FUNCTION_BLOCK "Conveyor_HMI_FB_1"   // FB 13, author

VAR_INPUT
   HMI_No : UInt;
   Sys_No : UInt;
   Zone : UInt;
END_VAR

VAR_IN_OUT
   Enable : Bool;
   Mode_Change : UInt;
   Transfer_To_ID : DInt;
   Transfer_From_ID : DInt;
   Pallet_Allignment : Bool;
   Enable(1) : Bool;
   Mode_Change(1) : UInt;
   Transfer_To_ID(1) : DInt;
   Transfer_From_ID(1) : DInt;
   Pallet_Allignment(1) : Bool;
END_VAR

VAR
   R_Charge_Cnv_Commands : R_TRIG;
   T_Reset_Charge : TON_TIME;
   ID : DInt;
   ID(1) : DInt;
   ID_Old : DInt;
   ID_Old(1) : DInt;
END_VAR

VAR_TEMP
   i : UInt;
   J : UInt;
   No_Light_Guard : Bool;
END_VAR

BEGIN
CNV_Selector_1(Sys_No := #Sys_No,
                 Zone:= #Zone,
                 CNV1_2_Selected := "CNV_HMI".CNV2_Selected[#HMI_No],
                 ID => #ID,
                 ID(1) => #"ID(1)");


REGION SEND/RECEIVE BUTTON
    IF NOT "Control_DB".VTD_Sys[#Sys_No].Running AND "Control_DB".VTD_Sys[#Sys_No].Current_Level <> 0 THEN
        IF "CNV_HMI".CNV2_Selected[#HMI_No] = 1 AND "HMI_DB".ScreenNo[#HMI_No] = 2 THEN
            //CNV 1
            IF "Control_DB".ECnv_Sys[#Sys_No].Cnv_Occupied AND NOT "Control_DB".LCnv_Sys[#Sys_No].Cnv_Level["Control_DB".VTD_Sys[#Sys_No].Current_Level].Cnv1.Cnv_Occupied AND
                NOT "Control_DB".ECnv_Sys[#Sys_No].Running AND NOT "Control_DB".LCnv_Sys[#Sys_No].Cnv_Level["Control_DB".VTD_Sys[#Sys_No].Current_Level].Cnv1.Running THEN
                "CNV_HMI".In_Out[#HMI_No] := TRUE;
            ELSIF NOT "Control_DB".ECnv_Sys[#Sys_No].Cnv_Occupied AND "Control_DB".LCnv_Sys[#Sys_No].Cnv_Level["Control_DB".VTD_Sys[#Sys_No].Current_Level].Cnv1.Cnv_Occupied AND
                NOT "Control_DB".ECnv_Sys[#Sys_No].Running AND NOT "Control_DB".LCnv_Sys[#Sys_No].Cnv_Level["Control_DB".VTD_Sys[#Sys_No].Current_Level].Cnv1.Running THEN
                "CNV_HMI".In_Out[#HMI_No] := FALSE;
            ELSE
                ;
            END_IF;
            //CNV 2
        ELSIF "CNV_HMI".CNV2_Selected[#HMI_No] = 2 AND "HMI_DB".ScreenNo[#HMI_No] = 2 THEN   //CNV 2
            IF "Control_DB".ECnv_Sys[#Sys_No].Cnv_Occupied AND NOT "Control_DB".LCnv_Sys[#Sys_No].Cnv_Level["Control_DB".VTD_Sys[#Sys_No].Current_Level].Cnv2.Cnv_Occupied AND
                NOT "Control_DB".ECnv_Sys[#Sys_No].Running AND NOT "Control_DB".LCnv_Sys[#Sys_No].Cnv_Level["Control_DB".VTD_Sys[#Sys_No].Current_Level].Cnv2.Running THEN
                "CNV_HMI".In_Out[#HMI_No] := TRUE;
            ELSIF NOT "Control_DB".ECnv_Sys[#Sys_No].Cnv_Occupied AND "Control_DB".LCnv_Sys[#Sys_No].Cnv_Level["Control_DB".VTD_Sys[#Sys_No].Current_Level].Cnv2.Cnv_Occupied AND
                NOT "Control_DB".ECnv_Sys[#Sys_No].Running AND NOT "Control_DB".LCnv_Sys[#Sys_No].Cnv_Level["Control_DB".VTD_Sys[#Sys_No].Current_Level].Cnv2.Running THEN
                "CNV_HMI".In_Out[#HMI_No] := FALSE;
            ELSE
                ;
            END_IF;
        END_IF;
    END_IF;
END_REGION ;

REGION Assign Conveyor 1
    REGION CHARGE DATA FROM THE CORRECT CONVEYOR
        //CHARGE DATA CHANGING CONVEYORS ID
        IF #ID <> #ID_Old THEN
            "CNV_HMI".Charge_Commands[#HMI_No] := TRUE;
            #ID_Old := #ID;
        END_IF;
        #R_Charge_Cnv_Commands();

        #R_Charge_Cnv_Commands(CLK := "CNV_HMI".Charge_Commands[#HMI_No]);

        //CHARGE ONCE THE COMMANDS
        IF "CNV_HMI".Charge_Commands[#Sys_No] THEN
            #Enable := "Control_DB".ECnv_Sys[#Sys_No].Instruction.Enable;
            #Mode_Change := "Control_DB".ECnv_Sys[#Sys_No].Instruction.Mode_Change;
            #Transfer_To_ID := "Control_DB".ECnv_Sys[#Sys_No].Instruction.Transfer_To_ID;
            #Transfer_From_ID := "Control_DB".ECnv_Sys[#Sys_No].Instruction.Transfer_From_ID;
            #Pallet_Allignment := "Control_DB".ECnv_Sys[#Sys_No].Instruction.Pallet_Allignment;
        END_IF;
    END_REGION

    REGION CHARGE DATA FROM HMI (AFTER CHARGE DATA)
        IF NOT "CNV_HMI".Charge_Commands[#HMI_No] AND NOT #R_Charge_Cnv_Commands.Q THEN
            CASE #ID OF
                    //SYSTEM 1
                120101:
                    Feed_ECNV_1(HMI_No := #HMI_No,
                                  HMI_Box:= #Zone,
                                  Overhang_Left:="CVTD1 OVERHANG LEFT",
                                  Overhang_Right:="CVTD1 OVERHANG RIGHT",
                                  Sys_No := #Sys_No,
                                  Safety_OK := "Remote_Panel_DB_1".Safety_OK);
                120201:
                    Feed_ECNV_1(HMI_No := #HMI_No,
                                  HMI_Box:= #Zone,
                                  Overhang_Left:="CVTD1 OVERHANG LEFT",
                                  Overhang_Right:="CVTD1 OVERHANG RIGHT",
                                  Sys_No := #Sys_No,
                                  Safety_OK := "Remote_Panel_DB_1".Safety_OK);
                120301:
                    Feed_ECNV_1(HMI_No := #HMI_No,
                                  HMI_Box:= #Zone,
                                  Overhang_Left:="CVTD1 OVERHANG LEFT",
                                  Overhang_Right:="CVTD1 OVERHANG RIGHT",
                                  Sys_No := #Sys_No,
                                  Safety_OK := "Remote_Panel_DB_1".Safety_OK);
                120401:
                    Feed_ECNV_1(HMI_No := #HMI_No,
                                  HMI_Box:= #Zone,
                                  Overhang_Left:="CVTD1 OVERHANG LEFT",
                                  Overhang_Right:="CVTD1 OVERHANG RIGHT",
                                  Sys_No := #Sys_No,
                                  Safety_OK := "Remote_Panel_DB_1".Safety_OK);
                120501:
                    Feed_ECNV_1(HMI_No := #HMI_No,
                                  HMI_Box:= #Zone,
                                  Overhang_Left:="CVTD1 OVERHANG LEFT",
                                  Overhang_Right:="CVTD1 OVERHANG RIGHT",
                                  Sys_No := #Sys_No,
                                  Safety_OK := "Remote_Panel_DB_1".Safety_OK);
                120601:
                    Feed_ECNV_1(HMI_No := #HMI_No,
                                  HMI_Box:= #Zone,
                                  Overhang_Left:="CVTD1 OVERHANG LEFT",
                                  Overhang_Right:="CVTD1 OVERHANG RIGHT",
                                  Sys_No := #Sys_No,
                                  Safety_OK := "Remote_Panel_DB_1".Safety_OK);
                120701:
                    Feed_ECNV_1(HMI_No := #HMI_No,
                                  HMI_Box:= #Zone,
                                  Overhang_Left:="CVTD1 OVERHANG LEFT",
                                  Overhang_Right:="CVTD1 OVERHANG RIGHT",
                                  Sys_No := #Sys_No,
                                  Safety_OK := "Remote_Panel_DB_1".Safety_OK);
                120801:
                    Feed_ECNV_1(HMI_No := #HMI_No,
                                  HMI_Box:= #Zone,
                                  Overhang_Left:="CVTD1 OVERHANG LEFT",
                                  Overhang_Right:="CVTD1 OVERHANG RIGHT",
                                  Sys_No := #Sys_No,
                                  Safety_OK := "Remote_Panel_DB_1".Safety_OK);

                    //SYSTEM 2
                120102:
                    Feed_ECNV_1(HMI_No := #HMI_No,
                                  HMI_Box:= #Zone,
                                  Overhang_Left:="CVTD2 OVERHANG LEFT",
                                  Overhang_Right:="CVTD2 OVERHANG RIGHT",
                                  Sys_No := 2,
                                  Safety_OK := "Remote_Panel_DB_2".Safety_OK);
                120202:
                    Feed_ECNV_1(HMI_No := #HMI_No,
                                  HMI_Box:= #Zone,
                                  Overhang_Left:="CVTD2 OVERHANG LEFT",
                                  Overhang_Right:="CVTD2 OVERHANG RIGHT",
                                  Sys_No := 2,
                                  Safety_OK := "Remote_Panel_DB_2".Safety_OK);
                120302:
                    Feed_ECNV_1(HMI_No := #HMI_No,
                                  HMI_Box:= #Zone,
                                  Overhang_Left:="CVTD2 OVERHANG LEFT",
                                  Overhang_Right:="CVTD2 OVERHANG RIGHT",
                                  Sys_No := 2,
                                  Safety_OK := "Remote_Panel_DB_2".Safety_OK);
                120402:
                    Feed_ECNV_1(HMI_No := #HMI_No,
                                  HMI_Box:= #Zone,
                                  Overhang_Left:="CVTD2 OVERHANG LEFT",
                                  Overhang_Right:="CVTD2 OVERHANG RIGHT",
                                  Sys_No := 2,
                                  Safety_OK := "Remote_Panel_DB_2".Safety_OK);
                120502:
                    Feed_ECNV_1(HMI_No := #HMI_No,
                                  HMI_Box:= #Zone,
                                  Overhang_Left:="CVTD2 OVERHANG LEFT",
                                  Overhang_Right:="CVTD2 OVERHANG RIGHT",
                                  Sys_No := 2,
                                  Safety_OK := "Remote_Panel_DB_2".Safety_OK);
                120602:
                    Feed_ECNV_1(HMI_No := #HMI_No,
                                  HMI_Box:= #Zone,
                                  Overhang_Left:="CVTD2 OVERHANG LEFT",
                                  Overhang_Right:="CVTD2 OVERHANG RIGHT",
                                  Sys_No := 2,
                                  Safety_OK := "Remote_Panel_DB_2".Safety_OK);
                120702:
                    Feed_ECNV_1(HMI_No := #HMI_No,
                                  HMI_Box:= #Zone,
                                  Overhang_Left:="CVTD2 OVERHANG LEFT",
                                  Overhang_Right:="CVTD2 OVERHANG RIGHT",
                                  Sys_No := 2,
                                  Safety_OK := "Remote_Panel_DB_2".Safety_OK);
                120802:
                    Feed_ECNV_1(HMI_No := #HMI_No,
                                  HMI_Box:= #Zone,
                                  Overhang_Left:="CVTD2 OVERHANG LEFT",
                                  Overhang_Right:="CVTD2 OVERHANG RIGHT",
                                  Sys_No := 2,
                                  Safety_OK := "Remote_Panel_DB_2".Safety_OK);

                    //SYSTEM 3
                120103:
                    Feed_ECNV_1(HMI_No := #HMI_No,
                                  HMI_Box:= #Zone,
                                  Overhang_Left:="CVTD3 OVERHANG LEFT",
                                  Overhang_Right:="CVTD3 OVERHANG RIGHT",
                                  Sys_No := 3,
                                  Safety_OK := "Remote_Panel_DB_3".Safety_OK);
                120203:
                    Feed_ECNV_1(HMI_No := #HMI_No,
                                  HMI_Box:= #Zone,
                                  Overhang_Left:="CVTD3 OVERHANG LEFT",
                                  Overhang_Right:="CVTD3 OVERHANG RIGHT",
                                  Sys_No := 3,
                                  Safety_OK := "Remote_Panel_DB_3".Safety_OK);
                120303:
                    Feed_ECNV_1(HMI_No := #HMI_No,
                                  HMI_Box:= #Zone,
                                  Overhang_Left:="CVTD3 OVERHANG LEFT",
                                  Overhang_Right:="CVTD3 OVERHANG RIGHT",
                                  Sys_No := 3,
                                  Safety_OK := "Remote_Panel_DB_3".Safety_OK);
                120403:
                    Feed_ECNV_1(HMI_No := #HMI_No,
                                  HMI_Box:= #Zone,
                                  Overhang_Left:="CVTD3 OVERHANG LEFT",
                                  Overhang_Right:="CVTD3 OVERHANG RIGHT",
                                  Sys_No := 3,
                                  Safety_OK := "Remote_Panel_DB_3".Safety_OK);
                120503:
                    Feed_ECNV_1(HMI_No := #HMI_No,
                                  HMI_Box:= #Zone,
                                  Overhang_Left:="CVTD3 OVERHANG LEFT",
                                  Overhang_Right:="CVTD3 OVERHANG RIGHT",
                                  Sys_No := 3,
                                  Safety_OK := "Remote_Panel_DB_3".Safety_OK);
                120603:
                    Feed_ECNV_1(HMI_No := #HMI_No,
                                  HMI_Box:= #Zone,
                                  Overhang_Left:="CVTD3 OVERHANG LEFT",
                                  Overhang_Right:="CVTD3 OVERHANG RIGHT",
                                  Sys_No := 3,
                                  Safety_OK := "Remote_Panel_DB_3".Safety_OK);
                120703:
                    Feed_ECNV_1(HMI_No := #HMI_No,
                                  HMI_Box:= #Zone,
                                  Overhang_Left:="CVTD3 OVERHANG LEFT",
                                  Overhang_Right:="CVTD3 OVERHANG RIGHT",
                                  Sys_No := 3,
                                  Safety_OK := "Remote_Panel_DB_3".Safety_OK);
                120803:
                    Feed_ECNV_1(HMI_No := #HMI_No,
                                  HMI_Box:= #Zone,
                                  Overhang_Left:="CVTD3 OVERHANG LEFT",
                                  Overhang_Right:="CVTD3 OVERHANG RIGHT",
                                  Sys_No := 3,
                                  Safety_OK := "Remote_Panel_DB_3".Safety_OK);

                    //SYSTEM 4
                120104:
                    Feed_ECNV_1(HMI_No := #HMI_No,
                                  HMI_Box:= #Zone,
                                  Overhang_Left:="CVTD4 OVERHANG LEFT",
                                  Overhang_Right:="CVTD4 OVERHANG RIGHT",
                                  Sys_No := 4,
                                  Safety_OK := "Remote_Panel_DB_4".Safety_OK);
                120204:
                    Feed_ECNV_1(HMI_No := #HMI_No,
                                  HMI_Box:= #Zone,
                                  Overhang_Left:="CVTD4 OVERHANG LEFT",
                                  Overhang_Right:="CVTD4 OVERHANG RIGHT",
                                  Sys_No := 4,
                                  Safety_OK := "Remote_Panel_DB_4".Safety_OK);
                120304:
                    Feed_ECNV_1(HMI_No := #HMI_No,
                                  HMI_Box:= #Zone,
                                  Overhang_Left:="CVTD4 OVERHANG LEFT",
                                  Overhang_Right:="CVTD4 OVERHANG RIGHT",
                                  Sys_No := 4,
                                  Safety_OK := "Remote_Panel_DB_4".Safety_OK);
                120404:
                    Feed_ECNV_1(HMI_No := #HMI_No,
                                  HMI_Box:= #Zone,
                                  Overhang_Left:="CVTD4 OVERHANG LEFT",
                                  Overhang_Right:="CVTD4 OVERHANG RIGHT",
                                  Sys_No := 4,
                                  Safety_OK := "Remote_Panel_DB_4".Safety_OK);
                120504:
                    Feed_ECNV_1(HMI_No := #HMI_No,
                                  HMI_Box:= #Zone,
                                  Overhang_Left:="CVTD4 OVERHANG LEFT",
                                  Overhang_Right:="CVTD4 OVERHANG RIGHT",
                                  Sys_No := 4,
                                  Safety_OK := "Remote_Panel_DB_4".Safety_OK);
                120604:
                    Feed_ECNV_1(HMI_No := #HMI_No,
                                  HMI_Box:= #Zone,
                                  Overhang_Left:="CVTD4 OVERHANG LEFT",
                                  Overhang_Right:="CVTD4 OVERHANG RIGHT",
                                  Sys_No := 4,
                                  Safety_OK := "Remote_Panel_DB_4".Safety_OK);
                120704:
                    Feed_ECNV_1(HMI_No := #HMI_No,
                                  HMI_Box:= #Zone,
                                  Overhang_Left:="CVTD4 OVERHANG LEFT",
                                  Overhang_Right:="CVTD4 OVERHANG RIGHT",
                                  Sys_No := 4,
                                  Safety_OK := "Remote_Panel_DB_4".Safety_OK);
                120804:
                    Feed_ECNV_1(HMI_No := #HMI_No,
                                  HMI_Box:= #Zone,
                                  Overhang_Left:="CVTD4 OVERHANG LEFT",
                                  Overhang_Right:="CVTD4 OVERHANG RIGHT",
                                  Sys_No := 4,
                                  Safety_OK := "Remote_Panel_DB_4".Safety_OK);

                    //SYSTEM 5
                120105:
                    Feed_ECNV_1(HMI_No := #HMI_No,
                                  HMI_Box:= #Zone,
                                  Overhang_Left:="CVTD5 OVERHANG LEFT",
                                  Overhang_Right:="CVTD5 OVERHANG RIGHT",
                                  Sys_No := 5,
                                  Safety_OK := "Remote_Panel_DB_5".Safety_OK);
                120205:
                    Feed_ECNV_1(HMI_No := #HMI_No,
                                  HMI_Box:= #Zone,
                                  Overhang_Left:="CVTD5 OVERHANG LEFT",
                                  Overhang_Right:="CVTD5 OVERHANG RIGHT",
                                  Sys_No := 5,
                                  Safety_OK := "Remote_Panel_DB_5".Safety_OK);
                120305:
                    Feed_ECNV_1(HMI_No := #HMI_No,
                                  HMI_Box:= #Zone,
                                  Overhang_Left:="CVTD5 OVERHANG LEFT",
                                  Overhang_Right:="CVTD5 OVERHANG RIGHT",
                                  Sys_No := 5,
                                  Safety_OK := "Remote_Panel_DB_5".Safety_OK);
                120405:
                    Feed_ECNV_1(HMI_No := #HMI_No,
                                  HMI_Box:= #Zone,
                                  Overhang_Left:="CVTD5 OVERHANG LEFT",
                                  Overhang_Right:="CVTD5 OVERHANG RIGHT",
                                  Sys_No := 5,
                                  Safety_OK := "Remote_Panel_DB_5".Safety_OK);
                120505:
                    Feed_ECNV_1(HMI_No := #HMI_No,
                                  HMI_Box:= #Zone,
                                  Overhang_Left:="CVTD5 OVERHANG LEFT",
                                  Overhang_Right:="CVTD5 OVERHANG RIGHT",
                                  Sys_No := 5,
                                  Safety_OK := "Remote_Panel_DB_5".Safety_OK);
                120605:
                    Feed_ECNV_1(HMI_No := #HMI_No,
                                  HMI_Box:= #Zone,
                                  Overhang_Left:="CVTD5 OVERHANG LEFT",
                                  Overhang_Right:="CVTD5 OVERHANG RIGHT",
                                  Sys_No := 5,
                                  Safety_OK := "Remote_Panel_DB_5".Safety_OK);
                120705:
                    Feed_ECNV_1(HMI_No := #HMI_No,
                                  HMI_Box:= #Zone,
                                  Overhang_Left:="CVTD5 OVERHANG LEFT",
                                  Overhang_Right:="CVTD5 OVERHANG RIGHT",
                                  Sys_No := 5,
                                  Safety_OK := "Remote_Panel_DB_5".Safety_OK);
                120805:
                    Feed_ECNV_1(HMI_No := #HMI_No,
                                  HMI_Box:= #Zone,
                                  Overhang_Left:="CVTD5 OVERHANG LEFT",
                                  Overhang_Right:="CVTD5 OVERHANG RIGHT",
                                  Sys_No := 5,
                                  Safety_OK := "Remote_Panel_DB_5".Safety_OK);
            END_CASE;
        END_IF;
    END_REGION
END_REGION

REGION Assign Conveyor 2
    REGION CHARGE DATA FROM THE CORRECT CONVEYOR
        //CHARGE DATA CHANGING CONVEYORS ID
        IF #"ID(1)" <> #"ID_Old(1)" THEN
            "CNV_HMI".Charge_Commands[#HMI_No] := TRUE;
            #"ID_Old(1)" := #"ID(1)";
        END_IF;
        #R_Charge_Cnv_Commands(CLK := "CNV_HMI".Charge_Commands[#HMI_No]);

        IF "CNV_HMI".Charge_Commands[#HMI_No] THEN
            CASE #"ID(1)" OF
                    //CNV 1 - SYSTEM 1
                100101:
                    #"Enable(1)" := "Control_DB".LCnv_Sys[#Sys_No].Cnv_Level[1].Cnv1.Instruction.Enable;
                    #"Mode_Change(1)" := "Control_DB".LCnv_Sys[#Sys_No].Cnv_Level[1].Cnv1.Instruction.Mode_Change;
                    #"Transfer_To_ID(1)" := "Control_DB".LCnv_Sys[#Sys_No].Cnv_Level[1].Cnv1.Instruction.Transfer_To_ID;
                    #"Transfer_From_ID(1)" := "Control_DB".LCnv_Sys[#Sys_No].Cnv_Level[1].Cnv1.Instruction.Transfer_From_ID;
                    #"Pallet_Allignment(1)" := "Control_DB".LCnv_Sys[#Sys_No].Cnv_Level[1].Cnv1.Instruction.Pallet_Allignment;
                100201:
                    "Enable_HMI(1)" := "Control_DB".LCnv_Sys[#Sys_No].Cnv_Level[2].Cnv1.Instruction.Enable;
                    "Mode_Change_HMI(1)" := "Control_DB".LCnv_Sys[#Sys_No].Cnv_Level[2].Cnv1.Instruction.Mode_Change;
                    "Transfer_To_ID_HMI(1)" := "Control_DB".LCnv_Sys[#Sys_No].Cnv_Level[2].Cnv1.Instruction.Transfer_To_ID;
                    "Transfer_From_ID_HMI(1)" := "Control_DB".LCnv_Sys[#Sys_No].Cnv_Level[2].Cnv1.Instruction.Transfer_From_ID;
                    "Pallet_Allignment_HMI(1)" := "Control_DB".LCnv_Sys[#Sys_No].Cnv_Level[2].Cnv1.Instruction.Pallet_Allignment;
                100301:
                    "Enable_HMI(1)" := "Control_DB".LCnv_Sys[#Sys_No].Cnv_Level[3].Cnv1.Instruction.Enable;
                    "Mode_Change_HMI(1)" := "Control_DB".LCnv_Sys[#Sys_No].Cnv_Level[3].Cnv1.Instruction.Mode_Change;
                    "Transfer_To_ID_HMI(1)" := "Control_DB".LCnv_Sys[#Sys_No].Cnv_Level[3].Cnv1.Instruction.Transfer_To_ID;
                    "Transfer_From_ID_HMI(1)" := "Control_DB".LCnv_Sys[#Sys_No].Cnv_Level[3].Cnv1.Instruction.Transfer_From_ID;
                    "Pallet_Allignment_HMI(1)" := "Control_DB".LCnv_Sys[#Sys_No].Cnv_Level[3].Cnv1.Instruction.Pallet_Allignment;
                100401:
                    "Enable_HMI(1)" := "Control_DB".LCnv_Sys[#Sys_No].Cnv_Level[4].Cnv1.Instruction.Enable;
                    "Mode_Change_HMI(1)" := "Control_DB".LCnv_Sys[#Sys_No].Cnv_Level[4].Cnv1.Instruction.Mode_Change;
                    "Transfer_To_ID_HMI(1)" := "Control_DB".LCnv_Sys[#Sys_No].Cnv_Level[4].Cnv1.Instruction.Transfer_To_ID;
                    "Transfer_From_ID_HMI(1)" := "Control_DB".LCnv_Sys[#Sys_No].Cnv_Level[4].Cnv1.Instruction.Transfer_From_ID;
                    "Pallet_Allignment_HMI(1)" := "Control_DB".LCnv_Sys[#Sys_No].Cnv_Level[4].Cnv1.Instruction.Pallet_Allignment;
                100501:
                    "Enable_HMI(1)" := "Control_DB".LCnv_Sys[#Sys_No].Cnv_Level[5].Cnv1.Instruction.Enable;
                    "Mode_Change_HMI(1)" := "Control_DB".LCnv_Sys[#Sys_No].Cnv_Level[5].Cnv1.Instruction.Mode_Change;
                    "Task_ID_HMI(1)" := "Control_DB".LCnv_Sys[#Sys_No].Cnv_Level[5].Cnv1.Instruction.Task_ID;
                    "Transfer_To_ID_HMI(1)" := "Control_DB".LCnv_Sys[#Sys_No].Cnv_Level[5].Cnv1.Instruction.Transfer_To_ID;
                    "Transfer_From_ID_HMI(1)" := "Control_DB".LCnv_Sys[#Sys_No].Cnv_Level[5].Cnv1.Instruction.Transfer_From_ID;
                    "Pallet_Allignment_HMI(1)" := "Control_DB".LCnv_Sys[#Sys_No].Cnv_Level[5].Cnv1.Instruction.Pallet_Allignment;
                100601:
                    "Enable_HMI(1)" := "Control_DB".LCnv_Sys[#Sys_No].Cnv_Level[6].Cnv1.Instruction.Enable;
                    "Mode_Change_HMI(1)" := "Control_DB".LCnv_Sys[#Sys_No].Cnv_Level[6].Cnv1.Instruction.Mode_Change;
                    "Task_ID_HMI(1)" := "Control_DB".LCnv_Sys[#Sys_No].Cnv_Level[6].Cnv1.Instruction.Task_ID;
                    "Transfer_To_ID_HMI(1)" := "Control_DB".LCnv_Sys[#Sys_No].Cnv_Level[6].Cnv1.Instruction.Transfer_To_ID;
                    "Transfer_From_ID_HMI(1)" := "Control_DB".LCnv_Sys[#Sys_No].Cnv_Level[6].Cnv1.Instruction.Transfer_From_ID;
                    "Pallet_Allignment_HMI(1)" := "Control_DB".LCnv_Sys[#Sys_No].Cnv_Level[6].Cnv1.Instruction.Pallet_Allignment;
                100701:
                    "Enable_HMI(1)" := "Control_DB".LCnv_Sys[#Sys_No].Cnv_Level[7].Cnv1.Instruction.Enable;
                    "Mode_Change_HMI(1)" := "Control_DB".LCnv_Sys[#Sys_No].Cnv_Level[7].Cnv1.Instruction.Mode_Change;
                    "Task_ID_HMI(1)" := "Control_DB".LCnv_Sys[#Sys_No].Cnv_Level[7].Cnv1.Instruction.Task_ID;
                    "Transfer_To_ID_HMI(1)" := "Control_DB".LCnv_Sys[#Sys_No].Cnv_Level[7].Cnv1.Instruction.Transfer_To_ID;
                    "Transfer_From_ID_HMI(1)" := "Control_DB".LCnv_Sys[#Sys_No].Cnv_Level[7].Cnv1.Instruction.Transfer_From_ID;
                    "Pallet_Allignment_HMI(1)" := "Control_DB".LCnv_Sys[#Sys_No].Cnv_Level[7].Cnv1.Instruction.Pallet_Allignment;
                100801:
                    "Enable_HMI(1)" := "Control_DB".LCnv_Sys[#Sys_No].Cnv_Level[8].Cnv1.Instruction.Enable;
                    "Mode_Change_HMI(1)" := "Control_DB".LCnv_Sys[#Sys_No].Cnv_Level[8].Cnv1.Instruction.Mode_Change;
                    "Task_ID_HMI(1)" := "Control_DB".LCnv_Sys[#Sys_No].Cnv_Level[8].Cnv1.Instruction.Task_ID;
                    "Transfer_To_ID_HMI(1)" := "Control_DB".LCnv_Sys[#Sys_No].Cnv_Level[8].Cnv1.Instruction.Transfer_To_ID;
                    "Transfer_From_ID_HMI(1)" := "Control_DB".LCnv_Sys[#Sys_No].Cnv_Level[8].Cnv1.Instruction.Transfer_From_ID;
                    "Pallet_Allignment_HMI(1)" := "Control_DB".LCnv_Sys[#Sys_No].Cnv_Level[8].Cnv1.Instruction.Pallet_Allignment;
                    //CNV 2 - SYSTEM 1
                110101:
                    "Enable_HMI(1)" := "Control_DB".LCnv_Sys[#Sys_No].Cnv_Level[1].Cnv2.Instruction.Enable;
                    "Mode_Change_HMI(1)" := "Control_DB".LCnv_Sys[#Sys_No].Cnv_Level[1].Cnv2.Instruction.Mode_Change;
                    "Task_ID_HMI(1)" := "Control_DB".LCnv_Sys[#Sys_No].Cnv_Level[1].Cnv2.Instruction.Task_ID;
                    "Transfer_To_ID_HMI(1)" := "Control_DB".LCnv_Sys[#Sys_No].Cnv_Level[1].Cnv2.Instruction.Transfer_To_ID;
                    "Transfer_From_ID_HMI(1)" := "Control_DB".LCnv_Sys[#Sys_No].Cnv_Level[1].Cnv2.Instruction.Transfer_From_ID;
                    "Pallet_Allignment_HMI(1)" := "Control_DB".LCnv_Sys[#Sys_No].Cnv_Level[1].Cnv2.Instruction.Pallet_Allignment;
                110201:
                    "Enable_HMI(1)" := "Control_DB".LCnv_Sys[#Sys_No].Cnv_Level[2].Cnv2.Instruction.Enable;
                    "Mode_Change_HMI(1)" := "Control_DB".LCnv_Sys[#Sys_No].Cnv_Level[2].Cnv2.Instruction.Mode_Change;
                    "Task_ID_HMI(1)" := "Control_DB".LCnv_Sys[#Sys_No].Cnv_Level[2].Cnv2.Instruction.Task_ID;
                    "Transfer_To_ID_HMI(1)" := "Control_DB".LCnv_Sys[#Sys_No].Cnv_Level[2].Cnv2.Instruction.Transfer_To_ID;
                    "Transfer_From_ID_HMI(1)" := "Control_DB".LCnv_Sys[#Sys_No].Cnv_Level[2].Cnv2.Instruction.Transfer_From_ID;
                    "Pallet_Allignment_HMI(1)" := "Control_DB".LCnv_Sys[#Sys_No].Cnv_Level[2].Cnv2.Instruction.Pallet_Allignment;
                110301:
                    "Enable_HMI(1)" := "Control_DB".LCnv_Sys[#Sys_No].Cnv_Level[3].Cnv2.Instruction.Enable;
                    "Mode_Change_HMI(1)" := "Control_DB".LCnv_Sys[#Sys_No].Cnv_Level[3].Cnv2.Instruction.Mode_Change;
                    "Task_ID_HMI(1)" := "Control_DB".LCnv_Sys[#Sys_No].Cnv_Level[3].Cnv2.Instruction.Task_ID;
                    "Transfer_To_ID_HMI(1)" := "Control_DB".LCnv_Sys[#Sys_No].Cnv_Level[3].Cnv2.Instruction.Transfer_To_ID;
                    "Transfer_From_ID_HMI(1)" := "Control_DB".LCnv_Sys[#Sys_No].Cnv_Level[3].Cnv2.Instruction.Transfer_From_ID;
                    "Pallet_Allignment_HMI(1)" := "Control_DB".LCnv_Sys[#Sys_No].Cnv_Level[3].Cnv2.Instruction.Pallet_Allignment;
                110401:
                    "Enable_HMI(1)" := "Control_DB".LCnv_Sys[#Sys_No].Cnv_Level[4].Cnv2.Instruction.Enable;
                    "Mode_Change_HMI(1)" := "Control_DB".LCnv_Sys[#Sys_No].Cnv_Level[4].Cnv2.Instruction.Mode_Change;
                    "Task_ID_HMI(1)" := "Control_DB".LCnv_Sys[#Sys_No].Cnv_Level[4].Cnv2.Instruction.Task_ID;
                    "Transfer_To_ID_HMI(1)" := "Control_DB".LCnv_Sys[#Sys_No].Cnv_Level[4].Cnv2.Instruction.Transfer_To_ID;
                    "Transfer_From_ID_HMI(1)" := "Control_DB".LCnv_Sys[#Sys_No].Cnv_Level[4].Cnv2.Instruction.Transfer_From_ID;
                    "Pallet_Allignment_HMI(1)" := "Control_DB".LCnv_Sys[#Sys_No].Cnv_Level[4].Cnv2.Instruction.Pallet_Allignment;
                110501:
                    "Enable_HMI(1)" := "Control_DB".LCnv_Sys[#Sys_No].Cnv_Level[5].Cnv2.Instruction.Enable;
                    "Mode_Change_HMI(1)" := "Control_DB".LCnv_Sys[#Sys_No].Cnv_Level[5].Cnv2.Instruction.Mode_Change;
                    "Task_ID_HMI(1)" := "Control_DB".LCnv_Sys[#Sys_No].Cnv_Level[5].Cnv2.Instruction.Task_ID;
                    "Transfer_To_ID_HMI(1)" := "Control_DB".LCnv_Sys[#Sys_No].Cnv_Level[5].Cnv2.Instruction.Transfer_To_ID;
                    "Transfer_From_ID_HMI(1)" := "Control_DB".LCnv_Sys[#Sys_No].Cnv_Level[5].Cnv2.Instruction.Transfer_From_ID;
                    "Pallet_Allignment_HMI(1)" := "Control_DB".LCnv_Sys[#Sys_No].Cnv_Level[5].Cnv2.Instruction.Pallet_Allignment;
                110601:
                    "Enable_HMI(1)" := "Control_DB".LCnv_Sys[#Sys_No].Cnv_Level[6].Cnv2.Instruction.Enable;
                    "Mode_Change_HMI(1)" := "Control_DB".LCnv_Sys[#Sys_No].Cnv_Level[6].Cnv2.Instruction.Mode_Change;
                    "Task_ID_HMI(1)" := "Control_DB".LCnv_Sys[#Sys_No].Cnv_Level[6].Cnv2.Instruction.Task_ID;
                    "Transfer_To_ID_HMI(1)" := "Control_DB".LCnv_Sys[#Sys_No].Cnv_Level[6].Cnv2.Instruction.Transfer_To_ID;
                    "Transfer_From_ID_HMI(1)" := "Control_DB".LCnv_Sys[#Sys_No].Cnv_Level[6].Cnv2.Instruction.Transfer_From_ID;
                    "Pallet_Allignment_HMI(1)" := "Control_DB".LCnv_Sys[#Sys_No].Cnv_Level[6].Cnv2.Instruction.Pallet_Allignment;
                110701:
                    "Enable_HMI(1)" := "Control_DB".LCnv_Sys[#Sys_No].Cnv_Level[7].Cnv2.Instruction.Enable;
                    "Mode_Change_HMI(1)" := "Control_DB".LCnv_Sys[#Sys_No].Cnv_Level[7].Cnv2.Instruction.Mode_Change;
                    "Task_ID_HMI(1)" := "Control_DB".LCnv_Sys[#Sys_No].Cnv_Level[7].Cnv2.Instruction.Task_ID;
                    "Transfer_To_ID_HMI(1)" := "Control_DB".LCnv_Sys[#Sys_No].Cnv_Level[7].Cnv2.Instruction.Transfer_To_ID;
                    "Transfer_From_ID_HMI(1)" := "Control_DB".LCnv_Sys[#Sys_No].Cnv_Level[7].Cnv2.Instruction.Transfer_From_ID;
                    "Pallet_Allignment_HMI(1)" := "Control_DB".LCnv_Sys[#Sys_No].Cnv_Level[7].Cnv2.Instruction.Pallet_Allignment;
                110801:
                    "Enable_HMI(1)" := "Control_DB".LCnv_Sys[#Sys_No].Cnv_Level[8].Cnv2.Instruction.Enable;
                    "Mode_Change_HMI(1)" := "Control_DB".LCnv_Sys[#Sys_No].Cnv_Level[8].Cnv2.Instruction.Mode_Change;
                    "Task_ID_HMI(1)" := "Control_DB".LCnv_Sys[#Sys_No].Cnv_Level[8].Cnv2.Instruction.Task_ID;
                    "Transfer_To_ID_HMI(1)" := "Control_DB".LCnv_Sys[#Sys_No].Cnv_Level[8].Cnv2.Instruction.Transfer_To_ID;
                    "Transfer_From_ID_HMI(1)" := "Control_DB".LCnv_Sys[#Sys_No].Cnv_Level[8].Cnv2.Instruction.Transfer_From_ID;
                    "Pallet_Allignment_HMI(1)" := "Control_DB".LCnv_Sys[#Sys_No].Cnv_Level[8].Cnv2.Instruction.Pallet_Allignment;
                    //CNV 1 - SYSTEM 2
                100102:
                    "Enable_HMI(1)" := "Control_DB".LCnv_Sys[2].Cnv_Level[1].Cnv1.Instruction.Enable;
                    "Mode_Change_HMI(1)" := "Control_DB".LCnv_Sys[2].Cnv_Level[1].Cnv1.Instruction.Mode_Change;
                    "Task_ID_HMI(1)" := "Control_DB".LCnv_Sys[2].Cnv_Level[1].Cnv1.Instruction.Task_ID;
                    "Transfer_To_ID_HMI(1)" := "Control_DB".LCnv_Sys[2].Cnv_Level[1].Cnv1.Instruction.Transfer_To_ID;
                    "Transfer_From_ID_HMI(1)" := "Control_DB".LCnv_Sys[2].Cnv_Level[1].Cnv1.Instruction.Transfer_From_ID;
                    "Pallet_Allignment_HMI(1)" := "Control_DB".LCnv_Sys[2].Cnv_Level[1].Cnv1.Instruction.Pallet_Allignment;
                100202:
                    "Enable_HMI(1)" := "Control_DB".LCnv_Sys[2].Cnv_Level[2].Cnv1.Instruction.Enable;
                    "Mode_Change_HMI(1)" := "Control_DB".LCnv_Sys[2].Cnv_Level[2].Cnv1.Instruction.Mode_Change;
                    "Task_ID_HMI(1)" := "Control_DB".LCnv_Sys[2].Cnv_Level[2].Cnv1.Instruction.Task_ID;
                    "Transfer_To_ID_HMI(1)" := "Control_DB".LCnv_Sys[2].Cnv_Level[2].Cnv1.Instruction.Transfer_To_ID;
                    "Transfer_From_ID_HMI(1)" := "Control_DB".LCnv_Sys[2].Cnv_Level[2].Cnv1.Instruction.Transfer_From_ID;
                    "Pallet_Allignment_HMI(1)" := "Control_DB".LCnv_Sys[2].Cnv_Level[2].Cnv1.Instruction.Pallet_Allignment;
                100302:
                    "Enable_HMI(1)" := "Control_DB".LCnv_Sys[2].Cnv_Level[3].Cnv1.Instruction.Enable;
                    "Mode_Change_HMI(1)" := "Control_DB".LCnv_Sys[2].Cnv_Level[3].Cnv1.Instruction.Mode_Change;
                    "Task_ID_HMI(1)" := "Control_DB".LCnv_Sys[2].Cnv_Level[3].Cnv1.Instruction.Task_ID;
                    "Transfer_To_ID_HMI(1)" := "Control_DB".LCnv_Sys[2].Cnv_Level[3].Cnv1.Instruction.Transfer_To_ID;
                    "Transfer_From_ID_HMI(1)" := "Control_DB".LCnv_Sys[2].Cnv_Level[3].Cnv1.Instruction.Transfer_From_ID;
                    "Pallet_Allignment_HMI(1)" := "Control_DB".LCnv_Sys[2].Cnv_Level[3].Cnv1.Instruction.Pallet_Allignment;
                100402:
                    "Enable_HMI(1)" := "Control_DB".LCnv_Sys[2].Cnv_Level[4].Cnv1.Instruction.Enable;
                    "Mode_Change_HMI(1)" := "Control_DB".LCnv_Sys[2].Cnv_Level[4].Cnv1.Instruction.Mode_Change;
                    "Task_ID_HMI(1)" := "Control_DB".LCnv_Sys[2].Cnv_Level[4].Cnv1.Instruction.Task_ID;
                    "Transfer_To_ID_HMI(1)" := "Control_DB".LCnv_Sys[2].Cnv_Level[4].Cnv1.Instruction.Transfer_To_ID;
                    "Transfer_From_ID_HMI(1)" := "Control_DB".LCnv_Sys[2].Cnv_Level[4].Cnv1.Instruction.Transfer_From_ID;
                    "Pallet_Allignment_HMI(1)" := "Control_DB".LCnv_Sys[2].Cnv_Level[4].Cnv1.Instruction.Pallet_Allignment;
                100502:
                    "Enable_HMI(1)" := "Control_DB".LCnv_Sys[2].Cnv_Level[5].Cnv1.Instruction.Enable;
                    "Mode_Change_HMI(1)" := "Control_DB".LCnv_Sys[2].Cnv_Level[5].Cnv1.Instruction.Mode_Change;
                    "Task_ID_HMI(1)" := "Control_DB".LCnv_Sys[2].Cnv_Level[5].Cnv1.Instruction.Task_ID;
                    "Transfer_To_ID_HMI(1)" := "Control_DB".LCnv_Sys[2].Cnv_Level[5].Cnv1.Instruction.Transfer_To_ID;
                    "Transfer_From_ID_HMI(1)" := "Control_DB".LCnv_Sys[2].Cnv_Level[5].Cnv1.Instruction.Transfer_From_ID;
                    "Pallet_Allignment_HMI(1)" := "Control_DB".LCnv_Sys[2].Cnv_Level[5].Cnv1.Instruction.Pallet_Allignment;
                100602:
                    "Enable_HMI(1)" := "Control_DB".LCnv_Sys[2].Cnv_Level[6].Cnv1.Instruction.Enable;
                    "Mode_Change_HMI(1)" := "Control_DB".LCnv_Sys[2].Cnv_Level[6].Cnv1.Instruction.Mode_Change;
                    "Task_ID_HMI(1)" := "Control_DB".LCnv_Sys[2].Cnv_Level[6].Cnv1.Instruction.Task_ID;
                    "Transfer_To_ID_HMI(1)" := "Control_DB".LCnv_Sys[2].Cnv_Level[6].Cnv1.Instruction.Transfer_To_ID;
                    "Transfer_From_ID_HMI(1)" := "Control_DB".LCnv_Sys[2].Cnv_Level[6].Cnv1.Instruction.Transfer_From_ID;
                    "Pallet_Allignment_HMI(1)" := "Control_DB".LCnv_Sys[2].Cnv_Level[6].Cnv1.Instruction.Pallet_Allignment;
                100702:
                    "Enable_HMI(1)" := "Control_DB".LCnv_Sys[2].Cnv_Level[7].Cnv1.Instruction.Enable;
                    "Mode_Change_HMI(1)" := "Control_DB".LCnv_Sys[2].Cnv_Level[7].Cnv1.Instruction.Mode_Change;
                    "Task_ID_HMI(1)" := "Control_DB".LCnv_Sys[2].Cnv_Level[7].Cnv1.Instruction.Task_ID;
                    "Transfer_To_ID_HMI(1)" := "Control_DB".LCnv_Sys[2].Cnv_Level[7].Cnv1.Instruction.Transfer_To_ID;
                    "Transfer_From_ID_HMI(1)" := "Control_DB".LCnv_Sys[2].Cnv_Level[7].Cnv1.Instruction.Transfer_From_ID;
                    "Pallet_Allignment_HMI(1)" := "Control_DB".LCnv_Sys[2].Cnv_Level[7].Cnv1.Instruction.Pallet_Allignment;
                100802:
                    "Enable_HMI(1)" := "Control_DB".LCnv_Sys[2].Cnv_Level[8].Cnv1.Instruction.Enable;
                    "Mode_Change_HMI(1)" := "Control_DB".LCnv_Sys[2].Cnv_Level[8].Cnv1.Instruction.Mode_Change;
                    "Task_ID_HMI(1)" := "Control_DB".LCnv_Sys[2].Cnv_Level[8].Cnv1.Instruction.Task_ID;
                    "Transfer_To_ID_HMI(1)" := "Control_DB".LCnv_Sys[2].Cnv_Level[8].Cnv1.Instruction.Transfer_To_ID;
                    "Transfer_From_ID_HMI(1)" := "Control_DB".LCnv_Sys[2].Cnv_Level[8].Cnv1.Instruction.Transfer_From_ID;
                    "Pallet_Allignment_HMI(1)" := "Control_DB".LCnv_Sys[2].Cnv_Level[8].Cnv1.Instruction.Pallet_Allignment;
                    //CNV 2 - SYSTEM 2
                110102:
                    "Enable_HMI(1)" := "Control_DB".LCnv_Sys[2].Cnv_Level[1].Cnv2.Instruction.Enable;
                    "Mode_Change_HMI(1)" := "Control_DB".LCnv_Sys[2].Cnv_Level[1].Cnv2.Instruction.Mode_Change;
                    "Task_ID_HMI(1)" := "Control_DB".LCnv_Sys[2].Cnv_Level[1].Cnv2.Instruction.Task_ID;
                    "Transfer_To_ID_HMI(1)" := "Control_DB".LCnv_Sys[2].Cnv_Level[1].Cnv2.Instruction.Transfer_To_ID;
                    "Transfer_From_ID_HMI(1)" := "Control_DB".LCnv_Sys[2].Cnv_Level[1].Cnv2.Instruction.Transfer_From_ID;
                    "Pallet_Allignment_HMI(1)" := "Control_DB".LCnv_Sys[2].Cnv_Level[1].Cnv2.Instruction.Pallet_Allignment;
                110202:
                    "Enable_HMI(1)" := "Control_DB".LCnv_Sys[2].Cnv_Level[2].Cnv2.Instruction.Enable;
                    "Mode_Change_HMI(1)" := "Control_DB".LCnv_Sys[2].Cnv_Level[2].Cnv2.Instruction.Mode_Change;
                    "Task_ID_HMI(1)" := "Control_DB".LCnv_Sys[2].Cnv_Level[2].Cnv2.Instruction.Task_ID;
                    "Transfer_To_ID_HMI(1)" := "Control_DB".LCnv_Sys[2].Cnv_Level[2].Cnv2.Instruction.Transfer_To_ID;
                    "Transfer_From_ID_HMI(1)" := "Control_DB".LCnv_Sys[2].Cnv_Level[2].Cnv2.Instruction.Transfer_From_ID;
                    "Pallet_Allignment_HMI(1)" := "Control_DB".LCnv_Sys[2].Cnv_Level[2].Cnv2.Instruction.Pallet_Allignment;
                110302:
                    "Enable_HMI(1)" := "Control_DB".LCnv_Sys[2].Cnv_Level[3].Cnv2.Instruction.Enable;
                    "Mode_Change_HMI(1)" := "Control_DB".LCnv_Sys[2].Cnv_Level[3].Cnv2.Instruction.Mode_Change;
                    "Task_ID_HMI(1)" := "Control_DB".LCnv_Sys[2].Cnv_Level[3].Cnv2.Instruction.Task_ID;
                    "Transfer_To_ID_HMI(1)" := "Control_DB".LCnv_Sys[2].Cnv_Level[3].Cnv2.Instruction.Transfer_To_ID;
                    "Transfer_From_ID_HMI(1)" := "Control_DB".LCnv_Sys[2].Cnv_Level[3].Cnv2.Instruction.Transfer_From_ID;
                    "Pallet_Allignment_HMI(1)" := "Control_DB".LCnv_Sys[2].Cnv_Level[3].Cnv2.Instruction.Pallet_Allignment;
                110402:
                    "Enable_HMI(1)" := "Control_DB".LCnv_Sys[2].Cnv_Level[4].Cnv2.Instruction.Enable;
                    "Mode_Change_HMI(1)" := "Control_DB".LCnv_Sys[2].Cnv_Level[4].Cnv2.Instruction.Mode_Change;
                    "Task_ID_HMI(1)" := "Control_DB".LCnv_Sys[2].Cnv_Level[4].Cnv2.Instruction.Task_ID;
                    "Transfer_To_ID_HMI(1)" := "Control_DB".LCnv_Sys[2].Cnv_Level[4].Cnv2.Instruction.Transfer_To_ID;
                    "Transfer_From_ID_HMI(1)" := "Control_DB".LCnv_Sys[2].Cnv_Level[4].Cnv2.Instruction.Transfer_From_ID;
                    "Pallet_Allignment_HMI(1)" := "Control_DB".LCnv_Sys[2].Cnv_Level[4].Cnv2.Instruction.Pallet_Allignment;
                110502:
                    "Enable_HMI(1)" := "Control_DB".LCnv_Sys[2].Cnv_Level[5].Cnv2.Instruction.Enable;
                    "Mode_Change_HMI(1)" := "Control_DB".LCnv_Sys[2].Cnv_Level[5].Cnv2.Instruction.Mode_Change;
                    "Task_ID_HMI(1)" := "Control_DB".LCnv_Sys[2].Cnv_Level[5].Cnv2.Instruction.Task_ID;
                    "Transfer_To_ID_HMI(1)" := "Control_DB".LCnv_Sys[2].Cnv_Level[5].Cnv2.Instruction.Transfer_To_ID;
                    "Transfer_From_ID_HMI(1)" := "Control_DB".LCnv_Sys[2].Cnv_Level[5].Cnv2.Instruction.Transfer_From_ID;
                    "Pallet_Allignment_HMI(1)" := "Control_DB".LCnv_Sys[2].Cnv_Level[5].Cnv2.Instruction.Pallet_Allignment;
                110602:
                    "Enable_HMI(1)" := "Control_DB".LCnv_Sys[2].Cnv_Level[6].Cnv2.Instruction.Enable;
                    "Mode_Change_HMI(1)" := "Control_DB".LCnv_Sys[2].Cnv_Level[6].Cnv2.Instruction.Mode_Change;
                    "Task_ID_HMI(1)" := "Control_DB".LCnv_Sys[2].Cnv_Level[6].Cnv2.Instruction.Task_ID;
                    "Transfer_To_ID_HMI(1)" := "Control_DB".LCnv_Sys[2].Cnv_Level[6].Cnv2.Instruction.Transfer_To_ID;
                    "Transfer_From_ID_HMI(1)" := "Control_DB".LCnv_Sys[2].Cnv_Level[6].Cnv2.Instruction.Transfer_From_ID;
                    "Pallet_Allignment_HMI(1)" := "Control_DB".LCnv_Sys[2].Cnv_Level[6].Cnv2.Instruction.Pallet_Allignment;
                110702:
                    "Enable_HMI(1)" := "Control_DB".LCnv_Sys[2].Cnv_Level[7].Cnv2.Instruction.Enable;
                    "Mode_Change_HMI(1)" := "Control_DB".LCnv_Sys[2].Cnv_Level[7].Cnv2.Instruction.Mode_Change;
                    "Task_ID_HMI(1)" := "Control_DB".LCnv_Sys[2].Cnv_Level[7].Cnv2.Instruction.Task_ID;
                    "Transfer_To_ID_HMI(1)" := "Control_DB".LCnv_Sys[2].Cnv_Level[7].Cnv2.Instruction.Transfer_To_ID;
                    "Transfer_From_ID_HMI(1)" := "Control_DB".LCnv_Sys[2].Cnv_Level[7].Cnv2.Instruction.Transfer_From_ID;
                    "Pallet_Allignment_HMI(1)" := "Control_DB".LCnv_Sys[2].Cnv_Level[7].Cnv2.Instruction.Pallet_Allignment;
                110802:
                    "Enable_HMI(1)" := "Control_DB".LCnv_Sys[2].Cnv_Level[8].Cnv2.Instruction.Enable;
                    "Mode_Change_HMI(1)" := "Control_DB".LCnv_Sys[2].Cnv_Level[8].Cnv2.Instruction.Mode_Change;
                    "Task_ID_HMI(1)" := "Control_DB".LCnv_Sys[2].Cnv_Level[8].Cnv2.Instruction.Task_ID;
                    "Transfer_To_ID_HMI(1)" := "Control_DB".LCnv_Sys[2].Cnv_Level[8].Cnv2.Instruction.Transfer_To_ID;
                    "Transfer_From_ID_HMI(1)" := "Control_DB".LCnv_Sys[2].Cnv_Level[8].Cnv2.Instruction.Transfer_From_ID;
                    "Pallet_Allignment_HMI(1)" := "Control_DB".LCnv_Sys[2].Cnv_Level[8].Cnv2.Instruction.Pallet_Allignment;
                    //CNV 1 - SYSTEM 3
                100103:
                    "Enable_HMI(1)" := "Control_DB".LCnv_Sys[3].Cnv_Level[1].Cnv1.Instruction.Enable;
                    "Mode_Change_HMI(1)" := "Control_DB".LCnv_Sys[3].Cnv_Level[1].Cnv1.Instruction.Mode_Change;
                    "Task_ID_HMI(1)" := "Control_DB".LCnv_Sys[3].Cnv_Level[1].Cnv1.Instruction.Task_ID;
                    "Transfer_To_ID_HMI(1)" := "Control_DB".LCnv_Sys[3].Cnv_Level[1].Cnv1.Instruction.Transfer_To_ID;
                    "Transfer_From_ID_HMI(1)" := "Control_DB".LCnv_Sys[3].Cnv_Level[1].Cnv1.Instruction.Transfer_From_ID;
                    "Pallet_Allignment_HMI(1)" := "Control_DB".LCnv_Sys[3].Cnv_Level[1].Cnv1.Instruction.Pallet_Allignment;
                100203:
                    "Enable_HMI(1)" := "Control_DB".LCnv_Sys[3].Cnv_Level[2].Cnv1.Instruction.Enable;
                    "Mode_Change_HMI(1)" := "Control_DB".LCnv_Sys[3].Cnv_Level[2].Cnv1.Instruction.Mode_Change;
                    "Task_ID_HMI(1)" := "Control_DB".LCnv_Sys[3].Cnv_Level[2].Cnv1.Instruction.Task_ID;
                    "Transfer_To_ID_HMI(1)" := "Control_DB".LCnv_Sys[3].Cnv_Level[2].Cnv1.Instruction.Transfer_To_ID;
                    "Transfer_From_ID_HMI(1)" := "Control_DB".LCnv_Sys[3].Cnv_Level[2].Cnv1.Instruction.Transfer_From_ID;
                    "Pallet_Allignment_HMI(1)" := "Control_DB".LCnv_Sys[3].Cnv_Level[2].Cnv1.Instruction.Pallet_Allignment;
                100303:
                    "Enable_HMI(1)" := "Control_DB".LCnv_Sys[3].Cnv_Level[3].Cnv1.Instruction.Enable;
                    "Mode_Change_HMI(1)" := "Control_DB".LCnv_Sys[3].Cnv_Level[3].Cnv1.Instruction.Mode_Change;
                    "Task_ID_HMI(1)" := "Control_DB".LCnv_Sys[3].Cnv_Level[3].Cnv1.Instruction.Task_ID;
                    "Transfer_To_ID_HMI(1)" := "Control_DB".LCnv_Sys[3].Cnv_Level[3].Cnv1.Instruction.Transfer_To_ID;
                    "Transfer_From_ID_HMI(1)" := "Control_DB".LCnv_Sys[3].Cnv_Level[3].Cnv1.Instruction.Transfer_From_ID;
                    "Pallet_Allignment_HMI(1)" := "Control_DB".LCnv_Sys[3].Cnv_Level[3].Cnv1.Instruction.Pallet_Allignment;
                100403:
                    "Enable_HMI(1)" := "Control_DB".LCnv_Sys[3].Cnv_Level[4].Cnv1.Instruction.Enable;
                    "Mode_Change_HMI(1)" := "Control_DB".LCnv_Sys[3].Cnv_Level[4].Cnv1.Instruction.Mode_Change;
                    "Task_ID_HMI(1)" := "Control_DB".LCnv_Sys[3].Cnv_Level[4].Cnv1.Instruction.Task_ID;
                    "Transfer_To_ID_HMI(1)" := "Control_DB".LCnv_Sys[3].Cnv_Level[4].Cnv1.Instruction.Transfer_To_ID;
                    "Transfer_From_ID_HMI(1)" := "Control_DB".LCnv_Sys[3].Cnv_Level[4].Cnv1.Instruction.Transfer_From_ID;
                    "Pallet_Allignment_HMI(1)" := "Control_DB".LCnv_Sys[3].Cnv_Level[4].Cnv1.Instruction.Pallet_Allignment;
                100503:
                    "Enable_HMI(1)" := "Control_DB".LCnv_Sys[3].Cnv_Level[5].Cnv1.Instruction.Enable;
                    "Mode_Change_HMI(1)" := "Control_DB".LCnv_Sys[3].Cnv_Level[5].Cnv1.Instruction.Mode_Change;
                    "Task_ID_HMI(1)" := "Control_DB".LCnv_Sys[3].Cnv_Level[5].Cnv1.Instruction.Task_ID;
                    "Transfer_To_ID_HMI(1)" := "Control_DB".LCnv_Sys[3].Cnv_Level[5].Cnv1.Instruction.Transfer_To_ID;
                    "Transfer_From_ID_HMI(1)" := "Control_DB".LCnv_Sys[3].Cnv_Level[5].Cnv1.Instruction.Transfer_From_ID;
                    "Pallet_Allignment_HMI(1)" := "Control_DB".LCnv_Sys[3].Cnv_Level[5].Cnv1.Instruction.Pallet_Allignment;
                100603:
                    "Enable_HMI(1)" := "Control_DB".LCnv_Sys[3].Cnv_Level[6].Cnv1.Instruction.Enable;
                    "Mode_Change_HMI(1)" := "Control_DB".LCnv_Sys[3].Cnv_Level[6].Cnv1.Instruction.Mode_Change;
                    "Task_ID_HMI(1)" := "Control_DB".LCnv_Sys[3].Cnv_Level[6].Cnv1.Instruction.Task_ID;
                    "Transfer_To_ID_HMI(1)" := "Control_DB".LCnv_Sys[3].Cnv_Level[6].Cnv1.Instruction.Transfer_To_ID;
                    "Transfer_From_ID_HMI(1)" := "Control_DB".LCnv_Sys[3].Cnv_Level[6].Cnv1.Instruction.Transfer_From_ID;
                    "Pallet_Allignment_HMI(1)" := "Control_DB".LCnv_Sys[3].Cnv_Level[6].Cnv1.Instruction.Pallet_Allignment;
                100703:
                    "Enable_HMI(1)" := "Control_DB".LCnv_Sys[3].Cnv_Level[7].Cnv1.Instruction.Enable;
                    "Mode_Change_HMI(1)" := "Control_DB".LCnv_Sys[3].Cnv_Level[7].Cnv1.Instruction.Mode_Change;
                    "Task_ID_HMI(1)" := "Control_DB".LCnv_Sys[3].Cnv_Level[7].Cnv1.Instruction.Task_ID;
                    "Transfer_To_ID_HMI(1)" := "Control_DB".LCnv_Sys[3].Cnv_Level[7].Cnv1.Instruction.Transfer_To_ID;
                    "Transfer_From_ID_HMI(1)" := "Control_DB".LCnv_Sys[3].Cnv_Level[7].Cnv1.Instruction.Transfer_From_ID;
                    "Pallet_Allignment_HMI(1)" := "Control_DB".LCnv_Sys[3].Cnv_Level[7].Cnv1.Instruction.Pallet_Allignment;
                100803:
                    "Enable_HMI(1)" := "Control_DB".LCnv_Sys[3].Cnv_Level[8].Cnv1.Instruction.Enable;
                    "Mode_Change_HMI(1)" := "Control_DB".LCnv_Sys[3].Cnv_Level[8].Cnv1.Instruction.Mode_Change;
                    "Task_ID_HMI(1)" := "Control_DB".LCnv_Sys[3].Cnv_Level[8].Cnv1.Instruction.Task_ID;
                    "Transfer_To_ID_HMI(1)" := "Control_DB".LCnv_Sys[3].Cnv_Level[8].Cnv1.Instruction.Transfer_To_ID;
                    "Transfer_From_ID_HMI(1)" := "Control_DB".LCnv_Sys[3].Cnv_Level[8].Cnv1.Instruction.Transfer_From_ID;
                    "Pallet_Allignment_HMI(1)" := "Control_DB".LCnv_Sys[3].Cnv_Level[8].Cnv1.Instruction.Pallet_Allignment;
                    //CNV 2 - SYSTEM 3
                110103:
                    "Enable_HMI(1)" := "Control_DB".LCnv_Sys[3].Cnv_Level[1].Cnv2.Instruction.Enable;
                    "Mode_Change_HMI(1)" := "Control_DB".LCnv_Sys[3].Cnv_Level[1].Cnv2.Instruction.Mode_Change;
                    "Task_ID_HMI(1)" := "Control_DB".LCnv_Sys[3].Cnv_Level[1].Cnv2.Instruction.Task_ID;
                    "Transfer_To_ID_HMI(1)" := "Control_DB".LCnv_Sys[3].Cnv_Level[1].Cnv2.Instruction.Transfer_To_ID;
                    "Transfer_From_ID_HMI(1)" := "Control_DB".LCnv_Sys[3].Cnv_Level[1].Cnv2.Instruction.Transfer_From_ID;
                    "Pallet_Allignment_HMI(1)" := "Control_DB".LCnv_Sys[3].Cnv_Level[1].Cnv2.Instruction.Pallet_Allignment;
                110203:
                    "Enable_HMI(1)" := "Control_DB".LCnv_Sys[3].Cnv_Level[2].Cnv2.Instruction.Enable;
                    "Mode_Change_HMI(1)" := "Control_DB".LCnv_Sys[3].Cnv_Level[2].Cnv2.Instruction.Mode_Change;
                    "Task_ID_HMI(1)" := "Control_DB".LCnv_Sys[3].Cnv_Level[2].Cnv2.Instruction.Task_ID;
                    "Transfer_To_ID_HMI(1)" := "Control_DB".LCnv_Sys[3].Cnv_Level[2].Cnv2.Instruction.Transfer_To_ID;
                    "Transfer_From_ID_HMI(1)" := "Control_DB".LCnv_Sys[3].Cnv_Level[2].Cnv2.Instruction.Transfer_From_ID;
                    "Pallet_Allignment_HMI(1)" := "Control_DB".LCnv_Sys[3].Cnv_Level[2].Cnv2.Instruction.Pallet_Allignment;
                110303:
                    "Enable_HMI(1)" := "Control_DB".LCnv_Sys[3].Cnv_Level[3].Cnv2.Instruction.Enable;
                    "Mode_Change_HMI(1)" := "Control_DB".LCnv_Sys[3].Cnv_Level[3].Cnv2.Instruction.Mode_Change;
                    "Task_ID_HMI(1)" := "Control_DB".LCnv_Sys[3].Cnv_Level[3].Cnv2.Instruction.Task_ID;
                    "Transfer_To_ID_HMI(1)" := "Control_DB".LCnv_Sys[3].Cnv_Level[3].Cnv2.Instruction.Transfer_To_ID;
                    "Transfer_From_ID_HMI(1)" := "Control_DB".LCnv_Sys[3].Cnv_Level[3].Cnv2.Instruction.Transfer_From_ID;
                    "Pallet_Allignment_HMI(1)" := "Control_DB".LCnv_Sys[3].Cnv_Level[3].Cnv2.Instruction.Pallet_Allignment;
                110403:
                    "Enable_HMI(1)" := "Control_DB".LCnv_Sys[3].Cnv_Level[4].Cnv2.Instruction.Enable;
                    "Mode_Change_HMI(1)" := "Control_DB".LCnv_Sys[3].Cnv_Level[4].Cnv2.Instruction.Mode_Change;
                    "Task_ID_HMI(1)" := "Control_DB".LCnv_Sys[3].Cnv_Level[4].Cnv2.Instruction.Task_ID;
                    "Transfer_To_ID_HMI(1)" := "Control_DB".LCnv_Sys[3].Cnv_Level[4].Cnv2.Instruction.Transfer_To_ID;
                    "Transfer_From_ID_HMI(1)" := "Control_DB".LCnv_Sys[3].Cnv_Level[4].Cnv2.Instruction.Transfer_From_ID;
                    "Pallet_Allignment_HMI(1)" := "Control_DB".LCnv_Sys[3].Cnv_Level[4].Cnv2.Instruction.Pallet_Allignment;
                110503:
                    "Enable_HMI(1)" := "Control_DB".LCnv_Sys[3].Cnv_Level[5].Cnv2.Instruction.Enable;
                    "Mode_Change_HMI(1)" := "Control_DB".LCnv_Sys[3].Cnv_Level[5].Cnv2.Instruction.Mode_Change;
                    "Task_ID_HMI(1)" := "Control_DB".LCnv_Sys[3].Cnv_Level[5].Cnv2.Instruction.Task_ID;
                    "Transfer_To_ID_HMI(1)" := "Control_DB".LCnv_Sys[3].Cnv_Level[5].Cnv2.Instruction.Transfer_To_ID;
                    "Transfer_From_ID_HMI(1)" := "Control_DB".LCnv_Sys[3].Cnv_Level[5].Cnv2.Instruction.Transfer_From_ID;
                    "Pallet_Allignment_HMI(1)" := "Control_DB".LCnv_Sys[3].Cnv_Level[5].Cnv2.Instruction.Pallet_Allignment;
                110603:
                    "Enable_HMI(1)" := "Control_DB".LCnv_Sys[3].Cnv_Level[6].Cnv2.Instruction.Enable;
                    "Mode_Change_HMI(1)" := "Control_DB".LCnv_Sys[3].Cnv_Level[6].Cnv2.Instruction.Mode_Change;
                    "Task_ID_HMI(1)" := "Control_DB".LCnv_Sys[3].Cnv_Level[6].Cnv2.Instruction.Task_ID;
                    "Transfer_To_ID_HMI(1)" := "Control_DB".LCnv_Sys[3].Cnv_Level[6].Cnv2.Instruction.Transfer_To_ID;
                    "Transfer_From_ID_HMI(1)" := "Control_DB".LCnv_Sys[3].Cnv_Level[6].Cnv2.Instruction.Transfer_From_ID;
                    "Pallet_Allignment_HMI(1)" := "Control_DB".LCnv_Sys[3].Cnv_Level[6].Cnv2.Instruction.Pallet_Allignment;
                110703:
                    "Enable_HMI(1)" := "Control_DB".LCnv_Sys[3].Cnv_Level[7].Cnv2.Instruction.Enable;
                    "Mode_Change_HMI(1)" := "Control_DB".LCnv_Sys[3].Cnv_Level[7].Cnv2.Instruction.Mode_Change;
                    "Task_ID_HMI(1)" := "Control_DB".LCnv_Sys[3].Cnv_Level[7].Cnv2.Instruction.Task_ID;
                    "Transfer_To_ID_HMI(1)" := "Control_DB".LCnv_Sys[3].Cnv_Level[7].Cnv2.Instruction.Transfer_To_ID;
                    "Transfer_From_ID_HMI(1)" := "Control_DB".LCnv_Sys[3].Cnv_Level[7].Cnv2.Instruction.Transfer_From_ID;
                    "Pallet_Allignment_HMI(1)" := "Control_DB".LCnv_Sys[3].Cnv_Level[7].Cnv2.Instruction.Pallet_Allignment;
                110803:
                    "Enable_HMI(1)" := "Control_DB".LCnv_Sys[3].Cnv_Level[8].Cnv2.Instruction.Enable;
                    "Mode_Change_HMI(1)" := "Control_DB".LCnv_Sys[3].Cnv_Level[8].Cnv2.Instruction.Mode_Change;
                    "Task_ID_HMI(1)" := "Control_DB".LCnv_Sys[3].Cnv_Level[8].Cnv2.Instruction.Task_ID;
                    "Transfer_To_ID_HMI(1)" := "Control_DB".LCnv_Sys[3].Cnv_Level[8].Cnv2.Instruction.Transfer_To_ID;
                    "Transfer_From_ID_HMI(1)" := "Control_DB".LCnv_Sys[3].Cnv_Level[8].Cnv2.Instruction.Transfer_From_ID;
                    "Pallet_Allignment_HMI(1)" := "Control_DB".LCnv_Sys[3].Cnv_Level[8].Cnv2.Instruction.Pallet_Allignment;
                    //CNV 2 - SYSTEM 4
                110104:
                    "Enable_HMI(1)" := "Control_DB".LCnv_Sys[4].Cnv_Level[1].Cnv2.Instruction.Enable;
                    "Mode_Change_HMI(1)" := "Control_DB".LCnv_Sys[4].Cnv_Level[1].Cnv2.Instruction.Mode_Change;
                    "Task_ID_HMI(1)" := "Control_DB".LCnv_Sys[4].Cnv_Level[1].Cnv2.Instruction.Task_ID;
                    "Transfer_To_ID_HMI(1)" := "Control_DB".LCnv_Sys[4].Cnv_Level[1].Cnv2.Instruction.Transfer_To_ID;
                    "Transfer_From_ID_HMI(1)" := "Control_DB".LCnv_Sys[4].Cnv_Level[1].Cnv2.Instruction.Transfer_From_ID;
                    "Pallet_Allignment_HMI(1)" := "Control_DB".LCnv_Sys[4].Cnv_Level[1].Cnv2.Instruction.Pallet_Allignment;
                110204:
                    "Enable_HMI(1)" := "Control_DB".LCnv_Sys[4].Cnv_Level[2].Cnv2.Instruction.Enable;
                    "Mode_Change_HMI(1)" := "Control_DB".LCnv_Sys[4].Cnv_Level[2].Cnv2.Instruction.Mode_Change;
                    "Task_ID_HMI(1)" := "Control_DB".LCnv_Sys[4].Cnv_Level[2].Cnv2.Instruction.Task_ID;
                    "Transfer_To_ID_HMI(1)" := "Control_DB".LCnv_Sys[4].Cnv_Level[2].Cnv2.Instruction.Transfer_To_ID;
                    "Transfer_From_ID_HMI(1)" := "Control_DB".LCnv_Sys[4].Cnv_Level[2].Cnv2.Instruction.Transfer_From_ID;
                    "Pallet_Allignment_HMI(1)" := "Control_DB".LCnv_Sys[4].Cnv_Level[2].Cnv2.Instruction.Pallet_Allignment;
                110304:
                    "Enable_HMI(1)" := "Control_DB".LCnv_Sys[4].Cnv_Level[3].Cnv2.Instruction.Enable;
                    "Mode_Change_HMI(1)" := "Control_DB".LCnv_Sys[4].Cnv_Level[3].Cnv2.Instruction.Mode_Change;
                    "Task_ID_HMI(1)" := "Control_DB".LCnv_Sys[4].Cnv_Level[3].Cnv2.Instruction.Task_ID;
                    "Transfer_To_ID_HMI(1)" := "Control_DB".LCnv_Sys[4].Cnv_Level[3].Cnv2.Instruction.Transfer_To_ID;
                    "Transfer_From_ID_HMI(1)" := "Control_DB".LCnv_Sys[4].Cnv_Level[3].Cnv2.Instruction.Transfer_From_ID;
                    "Pallet_Allignment_HMI(1)" := "Control_DB".LCnv_Sys[4].Cnv_Level[3].Cnv2.Instruction.Pallet_Allignment;
                110404:
                    "Enable_HMI(1)" := "Control_DB".LCnv_Sys[4].Cnv_Level[4].Cnv2.Instruction.Enable;
                    "Mode_Change_HMI(1)" := "Control_DB".LCnv_Sys[4].Cnv_Level[4].Cnv2.Instruction.Mode_Change;
                    "Task_ID_HMI(1)" := "Control_DB".LCnv_Sys[4].Cnv_Level[4].Cnv2.Instruction.Task_ID;
                    "Transfer_To_ID_HMI(1)" := "Control_DB".LCnv_Sys[4].Cnv_Level[4].Cnv2.Instruction.Transfer_To_ID;
                    "Transfer_From_ID_HMI(1)" := "Control_DB".LCnv_Sys[4].Cnv_Level[4].Cnv2.Instruction.Transfer_From_ID;
                    "Pallet_Allignment_HMI(1)" := "Control_DB".LCnv_Sys[4].Cnv_Level[4].Cnv2.Instruction.Pallet_Allignment;
                110504:
                    "Enable_HMI(1)" := "Control_DB".LCnv_Sys[4].Cnv_Level[5].Cnv2.Instruction.Enable;
                    "Mode_Change_HMI(1)" := "Control_DB".LCnv_Sys[4].Cnv_Level[5].Cnv2.Instruction.Mode_Change;
                    "Task_ID_HMI(1)" := "Control_DB".LCnv_Sys[4].Cnv_Level[5].Cnv2.Instruction.Task_ID;
                    "Transfer_To_ID_HMI(1)" := "Control_DB".LCnv_Sys[4].Cnv_Level[5].Cnv2.Instruction.Transfer_To_ID;
                    "Transfer_From_ID_HMI(1)" := "Control_DB".LCnv_Sys[4].Cnv_Level[5].Cnv2.Instruction.Transfer_From_ID;
                    "Pallet_Allignment_HMI(1)" := "Control_DB".LCnv_Sys[4].Cnv_Level[5].Cnv2.Instruction.Pallet_Allignment;
                110604:
                    "Enable_HMI(1)" := "Control_DB".LCnv_Sys[4].Cnv_Level[6].Cnv2.Instruction.Enable;
                    "Mode_Change_HMI(1)" := "Control_DB".LCnv_Sys[4].Cnv_Level[6].Cnv2.Instruction.Mode_Change;
                    "Task_ID_HMI(1)" := "Control_DB".LCnv_Sys[4].Cnv_Level[6].Cnv2.Instruction.Task_ID;
                    "Transfer_To_ID_HMI(1)" := "Control_DB".LCnv_Sys[4].Cnv_Level[6].Cnv2.Instruction.Transfer_To_ID;
                    "Transfer_From_ID_HMI(1)" := "Control_DB".LCnv_Sys[4].Cnv_Level[6].Cnv2.Instruction.Transfer_From_ID;
                    "Pallet_Allignment_HMI(1)" := "Control_DB".LCnv_Sys[4].Cnv_Level[6].Cnv2.Instruction.Pallet_Allignment;
                110704:
                    "Enable_HMI(1)" := "Control_DB".LCnv_Sys[4].Cnv_Level[7].Cnv2.Instruction.Enable;
                    "Mode_Change_HMI(1)" := "Control_DB".LCnv_Sys[4].Cnv_Level[7].Cnv2.Instruction.Mode_Change;
                    "Task_ID_HMI(1)" := "Control_DB".LCnv_Sys[4].Cnv_Level[7].Cnv2.Instruction.Task_ID;
                    "Transfer_To_ID_HMI(1)" := "Control_DB".LCnv_Sys[4].Cnv_Level[7].Cnv2.Instruction.Transfer_To_ID;
                    "Transfer_From_ID_HMI(1)" := "Control_DB".LCnv_Sys[4].Cnv_Level[7].Cnv2.Instruction.Transfer_From_ID;
                    "Pallet_Allignment_HMI(1)" := "Control_DB".LCnv_Sys[4].Cnv_Level[7].Cnv2.Instruction.Pallet_Allignment;
                110804:
                    "Enable_HMI(1)" := "Control_DB".LCnv_Sys[4].Cnv_Level[8].Cnv2.Instruction.Enable;
                    "Mode_Change_HMI(1)" := "Control_DB".LCnv_Sys[4].Cnv_Level[8].Cnv2.Instruction.Mode_Change;
                    "Task_ID_HMI(1)" := "Control_DB".LCnv_Sys[4].Cnv_Level[8].Cnv2.Instruction.Task_ID;
                    "Transfer_To_ID_HMI(1)" := "Control_DB".LCnv_Sys[4].Cnv_Level[8].Cnv2.Instruction.Transfer_To_ID;
                    "Transfer_From_ID_HMI(1)" := "Control_DB".LCnv_Sys[4].Cnv_Level[8].Cnv2.Instruction.Transfer_From_ID;
                    "Pallet_Allignment_HMI(1)" := "Control_DB".LCnv_Sys[4].Cnv_Level[8].Cnv2.Instruction.Pallet_Allignment;
                    //CNV 2 - SYSTEM 5
                110105:
                    "Enable_HMI(1)" := "Control_DB".LCnv_Sys[5].Cnv_Level[1].Cnv2.Instruction.Enable;
                    "Mode_Change_HMI(1)" := "Control_DB".LCnv_Sys[5].Cnv_Level[1].Cnv2.Instruction.Mode_Change;
                    "Task_ID_HMI(1)" := "Control_DB".LCnv_Sys[5].Cnv_Level[1].Cnv2.Instruction.Task_ID;
                    "Transfer_To_ID_HMI(1)" := "Control_DB".LCnv_Sys[5].Cnv_Level[1].Cnv2.Instruction.Transfer_To_ID;
                    "Transfer_From_ID_HMI(1)" := "Control_DB".LCnv_Sys[5].Cnv_Level[1].Cnv2.Instruction.Transfer_From_ID;
                    "Pallet_Allignment_HMI(1)" := "Control_DB".LCnv_Sys[5].Cnv_Level[1].Cnv2.Instruction.Pallet_Allignment;
                110205:
                    "Enable_HMI(1)" := "Control_DB".LCnv_Sys[5].Cnv_Level[2].Cnv2.Instruction.Enable;
                    "Mode_Change_HMI(1)" := "Control_DB".LCnv_Sys[5].Cnv_Level[2].Cnv2.Instruction.Mode_Change;
                    "Task_ID_HMI(1)" := "Control_DB".LCnv_Sys[5].Cnv_Level[2].Cnv2.Instruction.Task_ID;
                    "Transfer_To_ID_HMI(1)" := "Control_DB".LCnv_Sys[5].Cnv_Level[2].Cnv2.Instruction.Transfer_To_ID;
                    "Transfer_From_ID_HMI(1)" := "Control_DB".LCnv_Sys[5].Cnv_Level[2].Cnv2.Instruction.Transfer_From_ID;
                    "Pallet_Allignment_HMI(1)" := "Control_DB".LCnv_Sys[5].Cnv_Level[2].Cnv2.Instruction.Pallet_Allignment;
                110305:
                    "Enable_HMI(1)" := "Control_DB".LCnv_Sys[5].Cnv_Level[3].Cnv2.Instruction.Enable;
                    "Mode_Change_HMI(1)" := "Control_DB".LCnv_Sys[5].Cnv_Level[3].Cnv2.Instruction.Mode_Change;
                    "Task_ID_HMI(1)" := "Control_DB".LCnv_Sys[5].Cnv_Level[3].Cnv2.Instruction.Task_ID;
                    "Transfer_To_ID_HMI(1)" := "Control_DB".LCnv_Sys[5].Cnv_Level[3].Cnv2.Instruction.Transfer_To_ID;
                    "Transfer_From_ID_HMI(1)" := "Control_DB".LCnv_Sys[5].Cnv_Level[3].Cnv2.Instruction.Transfer_From_ID;
                    "Pallet_Allignment_HMI(1)" := "Control_DB".LCnv_Sys[5].Cnv_Level[3].Cnv2.Instruction.Pallet_Allignment;
                110405:
                    "Enable_HMI(1)" := "Control_DB".LCnv_Sys[5].Cnv_Level[4].Cnv2.Instruction.Enable;
                    "Mode_Change_HMI(1)" := "Control_DB".LCnv_Sys[5].Cnv_Level[4].Cnv2.Instruction.Mode_Change;
                    "Task_ID_HMI(1)" := "Control_DB".LCnv_Sys[5].Cnv_Level[4].Cnv2.Instruction.Task_ID;
                    "Transfer_To_ID_HMI(1)" := "Control_DB".LCnv_Sys[5].Cnv_Level[4].Cnv2.Instruction.Transfer_To_ID;
                    "Transfer_From_ID_HMI(1)" := "Control_DB".LCnv_Sys[5].Cnv_Level[4].Cnv2.Instruction.Transfer_From_ID;
                    "Pallet_Allignment_HMI(1)" := "Control_DB".LCnv_Sys[5].Cnv_Level[4].Cnv2.Instruction.Pallet_Allignment;
                110505:
                    "Enable_HMI(1)" := "Control_DB".LCnv_Sys[5].Cnv_Level[5].Cnv2.Instruction.Enable;
                    "Mode_Change_HMI(1)" := "Control_DB".LCnv_Sys[5].Cnv_Level[5].Cnv2.Instruction.Mode_Change;
                    "Task_ID_HMI(1)" := "Control_DB".LCnv_Sys[5].Cnv_Level[5].Cnv2.Instruction.Task_ID;
                    "Transfer_To_ID_HMI(1)" := "Control_DB".LCnv_Sys[5].Cnv_Level[5].Cnv2.Instruction.Transfer_To_ID;
                    "Transfer_From_ID_HMI(1)" := "Control_DB".LCnv_Sys[5].Cnv_Level[5].Cnv2.Instruction.Transfer_From_ID;
                    "Pallet_Allignment_HMI(1)" := "Control_DB".LCnv_Sys[5].Cnv_Level[5].Cnv2.Instruction.Pallet_Allignment;
                110605:
                    "Enable_HMI(1)" := "Control_DB".LCnv_Sys[5].Cnv_Level[6].Cnv2.Instruction.Enable;
                    "Mode_Change_HMI(1)" := "Control_DB".LCnv_Sys[5].Cnv_Level[6].Cnv2.Instruction.Mode_Change;
                    "Task_ID_HMI(1)" := "Control_DB".LCnv_Sys[5].Cnv_Level[6].Cnv2.Instruction.Task_ID;
                    "Transfer_To_ID_HMI(1)" := "Control_DB".LCnv_Sys[5].Cnv_Level[6].Cnv2.Instruction.Transfer_To_ID;
                    "Transfer_From_ID_HMI(1)" := "Control_DB".LCnv_Sys[5].Cnv_Level[6].Cnv2.Instruction.Transfer_From_ID;
                    "Pallet_Allignment_HMI(1)" := "Control_DB".LCnv_Sys[5].Cnv_Level[6].Cnv2.Instruction.Pallet_Allignment;
                110705:
                    "Enable_HMI(1)" := "Control_DB".LCnv_Sys[5].Cnv_Level[7].Cnv2.Instruction.Enable;
                    "Mode_Change_HMI(1)" := "Control_DB".LCnv_Sys[5].Cnv_Level[7].Cnv2.Instruction.Mode_Change;
                    "Task_ID_HMI(1)" := "Control_DB".LCnv_Sys[5].Cnv_Level[7].Cnv2.Instruction.Task_ID;
                    "Transfer_To_ID_HMI(1)" := "Control_DB".LCnv_Sys[5].Cnv_Level[7].Cnv2.Instruction.Transfer_To_ID;
                    "Transfer_From_ID_HMI(1)" := "Control_DB".LCnv_Sys[5].Cnv_Level[7].Cnv2.Instruction.Transfer_From_ID;
                    "Pallet_Allignment_HMI(1)" := "Control_DB".LCnv_Sys[5].Cnv_Level[7].Cnv2.Instruction.Pallet_Allignment;
                110805:
                    "Enable_HMI(1)" := "Control_DB".LCnv_Sys[5].Cnv_Level[8].Cnv2.Instruction.Enable;
                    "Mode_Change_HMI(1)" := "Control_DB".LCnv_Sys[5].Cnv_Level[8].Cnv2.Instruction.Mode_Change;
                    "Task_ID_HMI(1)" := "Control_DB".LCnv_Sys[5].Cnv_Level[8].Cnv2.Instruction.Task_ID;
                    "Transfer_To_ID_HMI(1)" := "Control_DB".LCnv_Sys[5].Cnv_Level[8].Cnv2.Instruction.Transfer_To_ID;
                    "Transfer_From_ID_HMI(1)" := "Control_DB".LCnv_Sys[5].Cnv_Level[8].Cnv2.Instruction.Transfer_From_ID;
                    "Pallet_Allignment_HMI(1)" := "Control_DB".LCnv_Sys[5].Cnv_Level[8].Cnv2.Instruction.Pallet_Allignment;
            END_CASE;
            "CNV_HMI".Charge_Commands[#HMI_No] := 0;
        END_IF;
    END_REGION

    REGION CHARGE DATA FROM HMI (AFTER CHARGE DATA)
        IF NOT "CNV_HMI".Charge_Commands[#HMI_No] AND NOT #R_Charge_Cnv_Commands.Q THEN
            CASE #"ID(1)" OF
                    //SYSTEM 1
                    //CNV 1
                100101:
                    "Feed_BCNV_Cnv1(1)_1"(HMI_No := #HMI_No,
                                          System_No := #Sys_No,
                                          Level := 1,
                                          Light_Guard_IO:="LIGHT GUARDS C1101 - CH1",
                                          Light_Guard_Bypass=>"Light_Guard_Bypass(1)");
                100201:
                    "Feed_BCNV_Cnv1(1)_1"(HMI_No := #HMI_No,
                                          System_No := #Sys_No,
                                          Level := 2,
                                          Light_Guard_IO:="LIGHT GUARDS C1101 - CH1",
                                          Light_Guard_Bypass=>"Light_Guard_Bypass(1)");
                100301:
                    "Feed_BCNV_Cnv1(1)_1"(HMI_No := #HMI_No,
                                          System_No := #Sys_No,
                                          Level := 3,
                                          Light_Guard_IO:="LIGHT GUARDS C1101 - CH1",
                                          Light_Guard_Bypass=>"Light_Guard_Bypass(1)");
                100401:
                    "Feed_BCNV_Cnv1(1)_1"(HMI_No := #HMI_No,
                                          System_No := #Sys_No,
                                          Level := 4,
                                          Light_Guard_IO:="LIGHT GUARDS C1101 - CH1",
                                          Light_Guard_Bypass=>"Light_Guard_Bypass(1)");
                100501:
                    "Feed_BCNV_Cnv1(1)_1"(HMI_No := #HMI_No,
                                          System_No := #Sys_No,
                                          Level := 5,
                                          Light_Guard_IO:="LIGHT GUARDS C1101 - CH1",
                                          Light_Guard_Bypass=>"Light_Guard_Bypass(1)");
                100601:
                    "Feed_BCNV_Cnv1(1)_1"(HMI_No := #HMI_No,
                                          System_No := #Sys_No,
                                          Level := 6,
                                          Light_Guard_IO:="LIGHT GUARDS C1101 - CH1",
                                          Light_Guard_Bypass=>"Light_Guard_Bypass(1)");
                100701:
                    "Feed_BCNV_Cnv1(1)_1"(HMI_No := #HMI_No,
                                          System_No := #Sys_No,
                                          Level := 7,
                                          Light_Guard_IO:="LIGHT GUARDS C1101 - CH1",
                                          Light_Guard_Bypass=>"Light_Guard_Bypass(1)");
                100801:
                    "Feed_BCNV_Cnv1(1)_1"(HMI_No := #HMI_No,
                                          System_No := #Sys_No,
                                          Level := 8,
                                          Light_Guard_IO:="LIGHT GUARDS C1101 - CH1",
                                          Light_Guard_Bypass=>"Light_Guard_Bypass(1)");
                    //CNV 2
                110101:
                    "Feed_BCNV_Cnv2(1)_1"(HMI_No := #HMI_No,
                                          System_No := #Sys_No,
                                          Level := 1,
                                          Light_Guard_IO:="LIGHT GUARDS C1201 - CH1",
                                          Light_Guard_Bypass=>"Light_Guard_Bypass(1)");
                110201:
                    "Feed_BCNV_Cnv2(1)_1"(HMI_No := #HMI_No,
                                          System_No := #Sys_No,
                                          Level := 2,
                                          Light_Guard_IO:="LIGHT GUARDS C1201 - CH1",
                                          Light_Guard_Bypass=>"Light_Guard_Bypass(1)");
                110301:
                    "Feed_BCNV_Cnv2(1)_1"(HMI_No := #HMI_No,
                                          System_No := #Sys_No,
                                          Level := 3,
                                          Light_Guard_IO:="LIGHT GUARDS C1201 - CH1",
                                          Light_Guard_Bypass=>"Light_Guard_Bypass(1)");
                110401:
                    "Feed_BCNV_Cnv2(1)_1"(HMI_No := #HMI_No,
                                          System_No := #Sys_No,
                                          Level := 4,
                                          Light_Guard_IO:="LIGHT GUARDS C1201 - CH1",
                                          Light_Guard_Bypass=>"Light_Guard_Bypass(1)");
                110501:
                    "Feed_BCNV_Cnv2(1)_1"(HMI_No := #HMI_No,
                                          System_No := #Sys_No,
                                          Level := 5,
                                          Light_Guard_IO:="LIGHT GUARDS C1201 - CH1",
                                          Light_Guard_Bypass=>"Light_Guard_Bypass(1)");
                110601:
                    "Feed_BCNV_Cnv2(1)_1"(HMI_No := #HMI_No,
                                          System_No := #Sys_No,
                                          Level := 6,
                                          Light_Guard_IO:="LIGHT GUARDS C1201 - CH1",
                                          Light_Guard_Bypass=>"Light_Guard_Bypass(1)");
                110701:
                    "Feed_BCNV_Cnv2(1)_1"(HMI_No := #HMI_No,
                                          System_No := #Sys_No,
                                          Level := 7,
                                          Light_Guard_IO:="LIGHT GUARDS C1201 - CH1",
                                          Light_Guard_Bypass=>"Light_Guard_Bypass(1)");
                110801:
                    "Feed_BCNV_Cnv2(1)_1"(HMI_No := #HMI_No,
                                          System_No := #Sys_No,
                                          Level := 8,
                                          Light_Guard_IO:="LIGHT GUARDS C1201 - CH1",
                                          Light_Guard_Bypass=>"Light_Guard_Bypass(1)");
                    //SYSTEM 2
                    //CNV 1
                100102:
                    "Feed_BCNV_Cnv1(1)_1"(HMI_No := #HMI_No,
                                          System_No := 2,
                                          Level := 1,
                                          Light_Guard_IO:="LIGHT GUARDS C2101 - CH1",
                                          Light_Guard_Bypass=>"Light_Guard_Bypass(2)");
                100202:
                    "Feed_BCNV_Cnv1(1)_1"(HMI_No := #HMI_No,
                                          System_No := 2,
                                          Level := 2,
                                          Light_Guard_IO:="LIGHT GUARDS C2101 - CH1",
                                          Light_Guard_Bypass=>"Light_Guard_Bypass(2)");
                100302:
                    "Feed_BCNV_Cnv1(1)_1"(HMI_No := #HMI_No,
                                          System_No := 2,
                                          Level := 3,
                                          Light_Guard_IO:="LIGHT GUARDS C2101 - CH1",
                                          Light_Guard_Bypass=>"Light_Guard_Bypass(2)");
                100402:
                    "Feed_BCNV_Cnv1(1)_1"(HMI_No := #HMI_No,
                                          System_No := 2,
                                          Level := 4,
                                          Light_Guard_IO:="LIGHT GUARDS C2101 - CH1",
                                          Light_Guard_Bypass=>"Light_Guard_Bypass(2)");
                100502:
                    "Feed_BCNV_Cnv1(1)_1"(HMI_No := #HMI_No,
                                          System_No := 2,
                                          Level := 5,
                                          Light_Guard_IO:="LIGHT GUARDS C2101 - CH1",
                                          Light_Guard_Bypass=>"Light_Guard_Bypass(2)");
                100602:
                    "Feed_BCNV_Cnv1(1)_1"(HMI_No := #HMI_No,
                                          System_No := 2,
                                          Level := 6,
                                          Light_Guard_IO:="LIGHT GUARDS C2101 - CH1",
                                          Light_Guard_Bypass=>"Light_Guard_Bypass(2)");
                100702:
                    "Feed_BCNV_Cnv1(1)_1"(HMI_No := #HMI_No,
                                          System_No := 2,
                                          Level := 7,
                                          Light_Guard_IO:="LIGHT GUARDS C2101 - CH1",
                                          Light_Guard_Bypass=>"Light_Guard_Bypass(2)");
                100802:
                    "Feed_BCNV_Cnv1(1)_1"(HMI_No := #HMI_No,
                                          System_No := 2,
                                          Level := 8,
                                          Light_Guard_IO:="LIGHT GUARDS C2101 - CH1",
                                          Light_Guard_Bypass=>"Light_Guard_Bypass(2)");
                    //CNV 2
                110102:
                    "Feed_BCNV_Cnv2(1)_1"(HMI_No := #HMI_No,
                                          System_No := 2,
                                          Level := 1,
                                          Light_Guard_IO:="LIGHT GUARDS C2201 - CH1",
                                          Light_Guard_Bypass=>"Light_Guard_Bypass(2)");
                110202:
                    "Feed_BCNV_Cnv2(1)_1"(HMI_No := #HMI_No,
                                          System_No := 2,
                                          Level := 2,
                                          Light_Guard_IO:="LIGHT GUARDS C2201 - CH1",
                                          Light_Guard_Bypass=>"Light_Guard_Bypass(2)");
                110302:
                    "Feed_BCNV_Cnv2(1)_1"(HMI_No := #HMI_No,
                                          System_No := 2,
                                          Level := 3,
                                          Light_Guard_IO:="LIGHT GUARDS C2201 - CH1",
                                          Light_Guard_Bypass=>"Light_Guard_Bypass(2)");
                110402:
                    "Feed_BCNV_Cnv2(1)_1"(HMI_No := #HMI_No,
                                          System_No := 2,
                                          Level := 4,
                                          Light_Guard_IO:="LIGHT GUARDS C2201 - CH1",
                                          Light_Guard_Bypass=>"Light_Guard_Bypass(2)");
                110502:
                    "Feed_BCNV_Cnv2(1)_1"(HMI_No := #HMI_No,
                                          System_No := 2,
                                          Level := 5,
                                          Light_Guard_IO:="LIGHT GUARDS C2201 - CH1",
                                          Light_Guard_Bypass=>"Light_Guard_Bypass(2)");
                110602:
                    "Feed_BCNV_Cnv2(1)_1"(HMI_No := #HMI_No,
                                          System_No := 2,
                                          Level := 6,
                                          Light_Guard_IO:="LIGHT GUARDS C2201 - CH1",
                                          Light_Guard_Bypass=>"Light_Guard_Bypass(2)");
                110702:
                    "Feed_BCNV_Cnv2(1)_1"(HMI_No := #HMI_No,
                                          System_No := 2,
                                          Level := 7,
                                          Light_Guard_IO:="LIGHT GUARDS C2201 - CH1",
                                          Light_Guard_Bypass=>"Light_Guard_Bypass(2)");
                110802:
                    "Feed_BCNV_Cnv2(1)_1"(HMI_No := #HMI_No,
                                          System_No := 2,
                                          Level := 8,
                                          Light_Guard_IO:="LIGHT GUARDS C2201 - CH1",
                                          Light_Guard_Bypass=>"Light_Guard_Bypass(2)");
                    //SYSTEM 3
                    //CNV 1
                100103:
                    "Feed_BCNV_Cnv1(1)_1"(HMI_No := #HMI_No,
                                          System_No := 3,
                                          Level := 1,
                                          Light_Guard_IO:="LIGHT GUARDS C3101 - CH1",
                                          Light_Guard_Bypass=>"Light_Guard_Bypass(3)");
                100203:
                    "Feed_BCNV_Cnv1(1)_1"(HMI_No := #HMI_No,
                                          System_No := 3,
                                          Level := 2,
                                          Light_Guard_IO:="LIGHT GUARDS C3101 - CH1",
                                          Light_Guard_Bypass=>"Light_Guard_Bypass(3)");
                100303:
                    "Feed_BCNV_Cnv1(1)_1"(HMI_No := #HMI_No,
                                          System_No := 3,
                                          Level := 3,
                                          Light_Guard_IO:="LIGHT GUARDS C3101 - CH1",
                                          Light_Guard_Bypass=>"Light_Guard_Bypass(3)");
                100403:
                    "Feed_BCNV_Cnv1(1)_1"(HMI_No := #HMI_No,
                                          System_No := 3,
                                          Level := 4,
                                          Light_Guard_IO:="LIGHT GUARDS C3101 - CH1",
                                          Light_Guard_Bypass=>"Light_Guard_Bypass(3)");
                100503:
                    "Feed_BCNV_Cnv1(1)_1"(HMI_No := #HMI_No,
                                          System_No := 3,
                                          Level := 5,
                                          Light_Guard_IO:="LIGHT GUARDS C3101 - CH1",
                                          Light_Guard_Bypass=>"Light_Guard_Bypass(3)");
                100603:
                    "Feed_BCNV_Cnv1(1)_1"(HMI_No := #HMI_No,
                                          System_No := 3,
                                          Level := 6,
                                          Light_Guard_IO:="LIGHT GUARDS C3101 - CH1",
                                          Light_Guard_Bypass=>"Light_Guard_Bypass(3)");
                100703:
                    "Feed_BCNV_Cnv1(1)_1"(HMI_No := #HMI_No,
                                          System_No := 3,
                                          Level := 7,
                                          Light_Guard_IO:="LIGHT GUARDS C3101 - CH1",
                                          Light_Guard_Bypass=>"Light_Guard_Bypass(3)");
                100803:
                    "Feed_BCNV_Cnv1(1)_1"(HMI_No := #HMI_No,
                                          System_No := 3,
                                          Level := 8,
                                          Light_Guard_IO:="LIGHT GUARDS C3101 - CH1",
                                          Light_Guard_Bypass=>"Light_Guard_Bypass(3)");
                    //CNV 2
                110103:
                    "Feed_BCNV_Cnv2(1)_1"(HMI_No := #HMI_No,
                                          System_No := 3,
                                          Level := 1,
                                          Light_Guard_IO:="LIGHT GUARDS C3201 - CH1",
                                          Light_Guard_Bypass=>"Light_Guard_Bypass(3)");
                110203:
                    "Feed_BCNV_Cnv2(1)_1"(HMI_No := #HMI_No,
                                          System_No := 3,
                                          Level := 2,
                                          Light_Guard_IO:="LIGHT GUARDS C3201 - CH1",
                                          Light_Guard_Bypass=>"Light_Guard_Bypass(3)");
                110303:
                    "Feed_BCNV_Cnv2(1)_1"(HMI_No := #HMI_No,
                                          System_No := 3,
                                          Level := 3,
                                          Light_Guard_IO:="LIGHT GUARDS C3201 - CH1",
                                          Light_Guard_Bypass=>"Light_Guard_Bypass(3)");
                110403:
                    "Feed_BCNV_Cnv2(1)_1"(HMI_No := #HMI_No,
                                          System_No := 3,
                                          Level := 4,
                                          Light_Guard_IO:="LIGHT GUARDS C3201 - CH1",
                                          Light_Guard_Bypass=>"Light_Guard_Bypass(3)");
                110503:
                    "Feed_BCNV_Cnv2(1)_1"(HMI_No := #HMI_No,
                                          System_No := 3,
                                          Level := 5,
                                          Light_Guard_IO:="LIGHT GUARDS C3201 - CH1",
                                          Light_Guard_Bypass=>"Light_Guard_Bypass(3)");
                110603:
                    "Feed_BCNV_Cnv2(1)_1"(HMI_No := #HMI_No,
                                          System_No := 3,
                                          Level := 6,
                                          Light_Guard_IO:="LIGHT GUARDS C3201 - CH1",
                                          Light_Guard_Bypass=>"Light_Guard_Bypass(3)");
                110703:
                    "Feed_BCNV_Cnv2(1)_1"(HMI_No := #HMI_No,
                                          System_No := 3,
                                          Level := 7,
                                          Light_Guard_IO:="LIGHT GUARDS C3201 - CH1",
                                          Light_Guard_Bypass=>"Light_Guard_Bypass(3)");
                110803:
                    "Feed_BCNV_Cnv2(1)_1"(HMI_No := #HMI_No,
                                          System_No := 3,
                                          Level := 8,
                                          Light_Guard_IO:="LIGHT GUARDS C3201 - CH1",
                                          Light_Guard_Bypass=>"Light_Guard_Bypass(3)");
                    //SYSTEM 4
                    //CNV 1
                100104:
                    "Feed_BCNV_Cnv2(1)_1"(HMI_No := #HMI_No,
                                          System_No := 4,
                                          Level := 1,
                                          Light_Guard_IO:=TRUE,
                                          Light_Guard_Bypass=>#No_Light_Guard);
                100204:
                    "Feed_BCNV_Cnv2(1)_1"(HMI_No := #HMI_No,
                                          System_No := 4,
                                          Level := 2,
                                          Light_Guard_IO:=TRUE,
                                          Light_Guard_Bypass=>#No_Light_Guard);
                100304:
                    "Feed_BCNV_Cnv2(1)_1"(HMI_No := #HMI_No,
                                          System_No := 4,
                                          Level := 3,
                                          Light_Guard_IO:=TRUE,
                                          Light_Guard_Bypass=>#No_Light_Guard);
                100404:
                    "Feed_BCNV_Cnv2(1)_1"(HMI_No := #HMI_No,
                                          System_No := 4,
                                          Level := 4,
                                          Light_Guard_IO:=TRUE,
                                          Light_Guard_Bypass=>#No_Light_Guard);
                100504:
                    "Feed_BCNV_Cnv2(1)_1"(HMI_No := #HMI_No,
                                          System_No := 4,
                                          Level := 5,
                                          Light_Guard_IO:=TRUE,
                                          Light_Guard_Bypass=>#No_Light_Guard);
                100604:
                    "Feed_BCNV_Cnv2(1)_1"(HMI_No := #HMI_No,
                                          System_No := 4,
                                          Level := 6,
                                          Light_Guard_IO:=TRUE,
                                          Light_Guard_Bypass=>#No_Light_Guard);
                100704:
                    "Feed_BCNV_Cnv2(1)_1"(HMI_No := #HMI_No,
                                          System_No := 4,
                                          Level := 7,
                                          Light_Guard_IO:=TRUE,
                                          Light_Guard_Bypass=>#No_Light_Guard);
                100804:
                    "Feed_BCNV_Cnv2(1)_1"(HMI_No := #HMI_No,
                                          System_No := 4,
                                          Level := 8,
                                          Light_Guard_IO:=TRUE,
                                          Light_Guard_Bypass=>#No_Light_Guard);
                    //SYSTEM 5
                    //CNV 1
                100105:
                    "Feed_BCNV_Cnv2(1)_1"(HMI_No := #HMI_No,
                                          System_No := 5,
                                          Level := 1,
                                          Light_Guard_IO:=TRUE,
                                          Light_Guard_Bypass=>#No_Light_Guard);
                100205:
                    "Feed_BCNV_Cnv2(1)_1"(HMI_No := #HMI_No,
                                          System_No := 5,
                                          Level := 2,
                                          Light_Guard_IO:=TRUE,
                                          Light_Guard_Bypass=>#No_Light_Guard);
                100305:
                    "Feed_BCNV_Cnv2(1)_1"(HMI_No := #HMI_No,
                                          System_No := 5,
                                          Level := 3,
                                          Light_Guard_IO:=TRUE,
                                          Light_Guard_Bypass=>#No_Light_Guard);
                100405:
                    "Feed_BCNV_Cnv2(1)_1"(HMI_No := #HMI_No,
                                          System_No := 5,
                                          Level := 4,
                                          Light_Guard_IO:=TRUE,
                                          Light_Guard_Bypass=>#No_Light_Guard);
                100505:
                    "Feed_BCNV_Cnv2(1)_1"(HMI_No := #HMI_No,
                                          System_No := 5,
                                          Level := 5,
                                          Light_Guard_IO:=TRUE,
                                          Light_Guard_Bypass=>#No_Light_Guard);
                100605:
                    "Feed_BCNV_Cnv2(1)_1"(HMI_No := #HMI_No,
                                          System_No := 5,
                                          Level := 6,
                                          Light_Guard_IO:=TRUE,
                                          Light_Guard_Bypass=>#No_Light_Guard);
                100705:
                    "Feed_BCNV_Cnv2(1)_1"(HMI_No := #HMI_No,
                                          System_No := 5,
                                          Level := 7,
                                          Light_Guard_IO:=TRUE,
                                          Light_Guard_Bypass=>#No_Light_Guard);
                100805:
                    "Feed_BCNV_Cnv2(1)_1"(HMI_No := #HMI_No,
                                          System_No := 5,
                                          Level := 8,
                                          Light_Guard_IO:=TRUE,
                                          Light_Guard_Bypass=>#No_Light_Guard);
            END_CASE;
        END_IF;
    END_REGION
END_REGION


//RESET CHARGE BITS
#T_Reset_Charge.TON(IN := "VTD_HMI".Charge_VTD[#HMI_No] OR "CNV_HMI".Charge_Cnv[#HMI_No] OR "VTD_HMI".Charge_VTD_Commands[#HMI_No] OR "CNV_HMI".Charge_Commands[#HMI_No],
                    PT := T#2S);

IF #T_Reset_Charge.Q THEN
    "VTD_HMI".Charge_VTD[#HMI_No] := FALSE;
    "CNV_HMI".Charge_Cnv[#HMI_No] := FALSE;
    "VTD_HMI".Charge_VTD_Commands[#HMI_No] := FALSE;
    "CNV_HMI".Charge_Commands[#HMI_No] := FALSE;
END_IF;

END_FUNCTION_BLOCK